(* IEC 61131-3 sources: daoli-st-library/DL_Process (part 30) *)

(* ---- FB_DL_DateCoderPosition.st ---- *)
(*==============================================================================
 * 组件名称 (Component)  : FB_DL_DateCoderPosition
 * 所属子库 (Sublibrary) : DL_Process
 * 当前版本 (Version)    : 1.0.0
 * 兼容性 (Platform)     : CODESYS 3.5+ / TwinCAT 3 / 汇川 InoProShop / 施耐德 Machine Expert
 *                         仅依赖 Standard.library（R_TRIG / ABS），零厂商私有库
 * 功能描述 (Function)   : 喷码日期位置偏移与缺失检测。检测触发沿按视觉检出
 *                         电平分派：未检出 → 缺失计数 + bMissing 锁存；检出
 *                         → 位置偏差 = 实测 - 期望，容差内 bPosOk，超差偏移
 *                         计数。判定结果锁存回放至下一触发沿（诊断资产）。
 *                         与 MarkPositionLatch（喷印位锁存）分工：本件是定
 *                         容差判偏移/缺失的诊断件。
 * 来源标签 (Origin)     : ROADMAP §21.4 R13 池（L907），自研 clean-room
 * 边界语义 (Boundary)   : ① 触发沿位置 NaN：按缺失域分派（视觉数据不可信 =
 *                         本拍无有效读码，归缺失语义安全侧）；
 *                         ② 容差/期望位置域闸 → 组态故障；
 *                         ③ 缺失/偏移计数 UDINT 独立成员（R190 归因唯一）；
 *                         ④ 状态锁存至下个触发沿（回放，不按当下输入重推断）。
 * 输出语义 (Fallback)   : 【R191】bEnable = FALSE → 判定出口冻结保持（诊断
 *                         资产）；eFault 相 → 冻结 + bError = TRUE。
 * 码位     (Codes)      : 按 R297 范式零 16# 码位硬编码；错误出口 BOOL+ENUM(eCause)。
 * 红线自检 (Redline)    : 7 项红线已自检：R1 零全局 ✓｜R2 零物理地址 ✓｜R3 纯 IEC ✓
 *                         R4 除零无涉/NaN 归缺失/组态闸 ✓｜R5 双语同行注释 ✓
 *                         R6 CASE 带 ELSE 兜底迁 eFault ✓｜R7 R_TRIG 段 0 无条件刷新 ✓
 * 验收向量 (Acceptance) : V1 期望 120.0、实测 121.4、容差 2.0 → 偏差 1.4，
 *                         bPosOk=TRUE；
 *                         V2 实测 124.0（偏差 4.0 超容差）→ nOffCnt+1，
 *                         bPosOk=FALSE；
 *                         V3 触发沿 bMarkPresent=FALSE → nMissCnt+1，
 *                         bMissing=TRUE。
 * 修订历史 (Revision)   : 2026-11-20  v1.0.0  R51 首版（批 3 · 序号 13）
 *==============================================================================*)
TYPE E_DL_DcpState :
(
    eIdle  := 0,                             (* 待使能 / Idle *)
    eInspect := 10,                          (* 检测运行 / Inspect run *)
    eFault := 90                             (* 故障锁存相 / Fault latched phase *)
);
END_TYPE

TYPE E_DL_DcpCause :
(
    eNone       := 0,                        (* 无故障成因 / No cause *)
    eCfgIllegal := 1,                        (* 组态非法：容差越域 / Illegal config *)
    ePhaseBad   := 2                         (* 非法相位兜底 / Illegal phase fallback *)
);
END_TYPE

FUNCTION_BLOCK FB_DL_DateCoderPosition
VAR_INPUT
    fMarkPos    : LREAL := 0.0;              (* 视觉测得喷码位置 [mm] / Measured mark position *)
    fMarkSp     : LREAL := 120.0;            (* 喷码期望位置，域 > 0 [mm] / Expected mark position *)
    fPosTol     : LREAL := 2.0;              (* 位置容差，域 > 0 [mm] / Position tolerance *)
    bMarkPresent: BOOL := FALSE;              (* 视觉检出电平 [-] / Vision present level *)
    bInspectTrig: BOOL := FALSE;             (* 检测触发电平（上升沿判定）[-] / Inspect trigger *)
    bEnable     : BOOL := TRUE;              (* 使能 [-] / Enable *)
    bReset      : BOOL := FALSE;             (* 复位命令，上升沿清全部 [-] / Reset command *)
END_VAR
VAR_OUTPUT
    fOffset     : LREAL;                     (* 位置偏差（实测 - 期望）[mm] / Position offset *)
    bPosOk      : BOOL;                      (* 位置合格判定（锁存回放）[-] / Position verdict *)
    bMissing    : BOOL;                      (* 喷码缺失锁存（下个触发沿或复位沿清）[-] / Missing latch *)
    nMissCnt    : UDINT;                     (* 缺失计数（独立成员，R190）[次] / Missing count *)
    nOffCnt     : UDINT;                     (* 偏移计数（独立成员，R190）[次] / Offset count *)
    nInspCnt    : UDINT;                     (* 累计检测次数 [次] / Inspect count *)
    eState      : E_DL_DcpState;             (* 状态出口 / State outlet *)
    eCause      : E_DL_DcpCause;             (* 故障成因出口 / Fault cause outlet *)
    bError      : BOOL;                      (* 故障锁存标志 [-] / Fault latch flag *)
END_VAR
VAR
    _eState   : E_DL_DcpState := E_DL_DcpState.eIdle;     (* 内部相位（CASE 唯一写入目标） / Internal phase *)
    _eCause   : E_DL_DcpCause := E_DL_DcpCause.eNone;     (* 故障成因锁存量 / Latched cause *)
    rtTrig    : R_TRIG;                      (* 触发沿实例，段 0 无条件调用 / Trigger edge instance *)
    rtReset   : R_TRIG;                      (* 复位沿实例，段 0 无条件调用 / Reset edge instance *)
    _fOff     : LREAL;                       (* 偏差派生量 [mm] / Offset derived *)
    _nMiss    : UDINT;                       (* 缺失计数锁存 [次] / Missing count latch *)
    _nOff     : UDINT;                       (* 偏移计数锁存 [次] / Offset count latch *)
    _nInsp    : UDINT;                       (* 检测计数锁存 [次] / Inspect count latch *)
    _bPosBad  : BOOL;                        (* 位置非有限当拍量 [-] / Non-finite position *)
    _bFault   : BOOL;                        (* 故障锁存位 / Latched fault bit *)
    _bCfgBad  : BOOL;                        (* 组态非法当拍量 / Illegal config this scan *)
END_VAR
VAR CONSTANT
    DL_DCP_EPS : LREAL := 1.0E-9;            (* 容差判零容差 [mm] / Tolerance epsilon *)
END_VAR

(* —— 段 0：当拍判据派生 + 沿实例无条件刷新（R228A） —— *)
_bCfgBad := (fPosTol <= DL_DCP_EPS) OR (fMarkSp <= 0.0);   (* 组态闸（R151 全引脚） / Config gate *)
rtTrig(CLK := bInspectTrig);                 (* 触发沿每拍必调 / Trigger edge every scan *)
rtReset(CLK := bReset);                      (* 复位沿每拍必调 / Reset edge every scan *)
_bPosBad := (fMarkPos <> fMarkPos) OR ((fMarkPos - fMarkPos) <> (fMarkPos - fMarkPos));   (* 位置 NaN 自反 + Inf 差判 / Non-finite position *)

(* —— 段 1：单拍量预清零（R107） —— *)
_fOff := 0.0;                                (* 偏差预清（判定拍内派生，R285） / Offset preset *)
bPosOk := FALSE;                             (* 判定预清（锁存拍内覆盖） / Verdict preset *)

(* —— 段 2：复位沿处理（作用域：清故障 + 清计数 + 清判定锁存 + 清出口 + 迁 eIdle，R283 逐项声明） —— *)
IF rtReset.Q THEN
    _bFault := FALSE;                        (* 清故障锁存 / Clear fault *)
    _eCause := E_DL_DcpCause.eNone;          (* 清成因 / Clear cause *)
    _nMiss := 0;                             (* 清缺失计数 / Clear miss count *)
    _nOff := 0;                              (* 清偏移计数 / Clear offset count *)
    _nInsp := 0;                             (* 清检测计数 / Clear inspect count *)
    bMissing := FALSE;                       (* 清缺失锁存（复位沿清除路径） / Clear missing latch *)
    bPosOk := FALSE;                         (* 清判定出口 / Clear verdict outlet *)
    fOffset := 0.0;                          (* 清偏差出口 / Clear offset outlet *)
    _eState := E_DL_DcpState.eIdle;          (* 迁待机相 / Back to idle *)
END_IF

(* —— 段 3：组态闸故障锁存（R45 配对；锁存至复位沿，R189） —— *)
IF _bCfgBad AND NOT _bFault THEN
    _bFault := TRUE;                         (* 锁存故障位 / Latch fault *)
    _eCause := E_DL_DcpCause.eCfgIllegal;    (* 成因：组态非法 / Cause: illegal config *)
    _eState := E_DL_DcpState.eFault;         (* 同步迁故障相 / Migrate to fault *)
END_IF

(* —— 段 4：CASE 主状态机（ELSE 兜底迁 eFault，红线 6） —— *)
CASE _eState OF
    E_DL_DcpState.eIdle:                     (* 待机相 / Idle *)
        IF bEnable AND NOT _bFault THEN
            _eState := E_DL_DcpState.eInspect;   (* 进入检测 / Enter inspect *)
        END_IF
    E_DL_DcpState.eInspect:                  (* 检测相：触发沿分派判定 / Inspect *)
        IF NOT bEnable THEN
            _eState := E_DL_DcpState.eIdle;  (* 失能回待机 / Back to idle *)
        ELSIF rtTrig.Q THEN                  (* 触发沿执行 / On trigger edge *)
            _nInsp := _nInsp + 1;            (* 检测计数（UDINT 回绕工程安全） / Count inspect *)
            IF (NOT bMarkPresent) OR _bPosBad THEN   (* 未检出或位置坏值：归缺失域（边界①安全侧） / Missing domain *)
                _nMiss := _nMiss + 1;        (* 缺失计数（独立成员） / Count missing *)
                bMissing := TRUE;            (* 缺失锁存（下个沿或复位清，边界④） / Latch missing *)
                bPosOk := FALSE;             (* 判定回放刷新 / Verdict replay *)
            ELSE
                _fOff := fMarkPos - fMarkSp; (* 偏差派生（减法无除零） / Offset derive *)
                fOffset := _fOff;            (* 偏差出口刷新 / Offset outlet *)
                IF ABS(_fOff) <= fPosTol THEN
                    bPosOk := TRUE;          (* 容差内合格 / In tolerance *)
                    bMissing := FALSE;       (* 检出合格拍清缺失锁存（触发沿清除路径，边界④） / Clear missing on pass *)
                ELSE
                    _nOff := _nOff + 1;      (* 偏移计数（独立成员） / Count offset *)
                    bPosOk := FALSE;         (* 超差不合格 / Out of tolerance *)
                END_IF
            END_IF
        END_IF                               (* 非触发拍：状态锁存回放（边界④） / Replay between edges *)
    E_DL_DcpState.eFault:                    (* 故障相：冻结保持，仅复位沿出 / Fault *)
        ;                                    (* 锁存回放（R28） / Replay from latch *)
    ELSE                                     (* 非法相位兜底迁安全态 / Illegal phase fallback *)
        _eState := E_DL_DcpState.eFault;     (* 迁故障相 / To fault *)
        _bFault := TRUE;                     (* 同步锁存 / Latch *)
        _eCause := E_DL_DcpCause.ePhaseBad;  (* 成因：非法相位 / Cause: illegal phase *)
END_CASE

(* —— 段 5：出口映射（bError/eState 同源，R191） —— *)
nMissCnt := _nMiss;                          (* 缺失计数出口 / Miss outlet *)
nOffCnt := _nOff;                            (* 偏移计数出口 / Offset outlet *)
nInspCnt := _nInsp;                          (* 检测计数出口 / Inspect outlet *)
bError := _bFault;                           (* 故障标志镜像 / Fault flag mirror *)
eState := _eState;                           (* 状态出口 / State outlet *)
eCause := _eCause;                           (* 成因出口 / Cause outlet *)
END_FUNCTION_BLOCK

(* ---- FB_DL_DesiccantRegenSeq.st ---- *)
(*
  组件名 Component   : FB_DL_DesiccantRegenSeq
  子库 Sublibrary    : DL_Process
  版本 Version       : 1.0.0
  兼容性 Platform    : CODESYS 3.5 / TwinCAT 3 / 汇川 InoProShop / Machine Expert（仅 Standard.library）
  功能 Function      : 干燥剂吸附塔再生顺控（ISA-88 相语义最小子集）：
                       1) 四相顺控：吸附（eAdsorb）→ 再生（eRegen）→ 吹冷（eCool）→
                       切换驻留（eSwitchDwell）→ 回吸附，吸附时长由 tAdsorbDur 承载；
                       2) 塔间轮换：A/B 双塔，eSwitchDwell 相完成阀组切换并翻转
                       bTowerAActive/bTowerBActive（切换指令单点出口）；
                       3) 再生温度曲线监视：再生相内再生温度须在
                       [fRegenTempLoC, fRegenTempHiC] 曲线带内，越带持续 tTempDevTo
                       → 故障锁存；
                       4) 各相计时独立 TON 实例（禁跨相复用，R228A）。
  边界 Boundary      : ① 本件只出阀组/加热指令与塔选通，不写物理 IO；
                       ② 吹冷相退出双条件：吹冷计时到 或 出口温度低于 fCoolEndC
                       （事件达成 + 前置消失双路径）；再生许可不满足时吸附相驻留等待；
                       ③ 故障锁存解除唯一路径 = bReset 上升沿（输入引脚，恒可达）；
                       ④ 无全局变量引用、无外部变量声明、无物理地址寻址。
  依赖 Depends       : Standard.library（R_TRIG / TON）
  溯源 Origin        : 道莅自研 clean-room（参考 t2-8-isa88 相语义分类与参数域，
                       零代码行复制）
  码位 Code          : 16#06_0_BE（Process 段 0006，B 子带 BE 格）
  码表 Error codes（本件格 06_0_BE，单轨子道：故障 0x02BE / 信息 0x01BE）:
    16#0006_02BE 故障级：再生顺控故障总码（再生温度越带 / 切换超时 / 组态非法 /
                 输入非有限），锁存至复位
    16#0006_01BE 信息级：塔切换完成沿（eSwitchDwell → eAdsorb 迁移拍）
  修订历史 Revision  :
    2026-11-19  v1.0.0  R44 首版（批次 3 · 序号 15）
*)

TYPE E_DL_DrsPhase :
(
    eIdle        := 0,   // 空闲：未使能 / Idle, not enabled
    eAdsorb      := 10,  // 吸附：当前塔吸附运行 / Adsorbing on active tower
    eRegen       := 20,  // 再生：离线塔再生加热 / Regenerating offline tower
    eCool        := 30,  // 吹冷：再生塔吹冷 / Cooling regenerated tower
    eSwitchDwell := 40,  // 切换：塔间阀组切换驻留 / Switching towers dwell
    eFault       := 90   // 故障：总码锁存 / Fault, latched
);
END_TYPE

FUNCTION_BLOCK FB_DL_DesiccantRegenSeq
VAR_INPUT
    bEnable      : BOOL;                   // 使能（电平）[-] / Enable
    bReset       : BOOL;                   // 上升沿清故障锁存 [-] / Reset edge
    bRegenPermissive: BOOL;                // 再生许可（电平）[-] / Regen permissive
    fRegenTempC  : REAL;                   // 再生温度 [摄氏度] / Regen temperature
    fCoolOutTempC: REAL;                   // 吹冷出口温度 [摄氏度] / Cooling outlet temperature
    tAdsorbDur   : TIME := T#8H;           // 吸附时长 [毫秒] / Adsorption duration
    tRegenDur    : TIME := T#4H;           // 再生时长 [毫秒] / Regen duration
    tCoolMaxDur  : TIME := T#2H;           // 吹冷最大时长 [毫秒] / Cooling max duration
    tSwitchDur   : TIME := T#60S;          // 切换驻留 [毫秒] / Switch dwell
    fRegenTempLoC: REAL := 120.0;          // 再生温度带下限 [摄氏度] / Regen band floor
    fRegenTempHiC: REAL := 200.0;          // 再生温度带上限 [摄氏度] / Regen band ceiling
    fCoolEndC    : REAL := 45.0;           // 吹冷结束温度 [摄氏度] / Cooling end temperature
    tTempDevTo   : TIME := T#30S;          // 温度越带确认窗 [毫秒] / Temperature deviation timeout
END_VAR
VAR_OUTPUT
    bTowerAActive: BOOL;                   // A 塔吸附选通 [-] / Tower A active
    bTowerBActive: BOOL;                   // B 塔吸附选通 [-] / Tower B active
    bRegenHeatCmd: BOOL;                   // 再生加热指令 [-] / Regen heat command
    bRegenCoolCmd: BOOL;                   // 吹冷指令 [-] / Regen cool command
    bSwitchCmd   : BOOL;                   // 塔切换指令（驻留相电平）[-] / Tower switch command
    ePhase       : E_DL_DrsPhase;          // 相位出口，段尾单点映射 / Phase outlet
    bError       : BOOL;                   // 故障锁存标志 [-] / Fault latch flag
    uErrId       : UDINT;                  // 事件码，0 = 无事件 / Event code
END_VAR
VAR
    rtReset   : R_TRIG;                    // 复位沿实例，段 0 无条件刷新 / Reset edge
    tonAdsorb : TON;                       // 吸附计时（独立实例） / Adsorption timer
    tonRegen  : TON;                       // 再生计时（独立实例） / Regen timer
    tonCoolMax: TON;                       // 吹冷最大计时（独立实例） / Cooling max timer
    tonSwitch : TON;                       // 切换驻留计时（独立实例） / Switch dwell timer
    tonTempDevTo: TON;                     // 温度越带确认（专用超时件命名） / Temp deviation timeout
    _ePhase   : E_DL_DrsPhase := E_DL_DrsPhase.eIdle;  // 内部相位（CASE 唯一写入目标）/ Internal phase
    _bTowerA  : BOOL := TRUE;              // 内部塔选（TRUE = A 塔吸附）/ Internal tower select
    _bFault   : BOOL;                      // 故障锁存位（锁存量） / Latched fault bit
    _uFault   : UDINT;                     // 故障码锁存（锁存量） / Latched fault code
    _bCfgBad  : BOOL;                      // 组态非法当拍量 [-] / Config illegal flag
    _bNonFin  : BOOL;                      // 输入非有限当拍量 [-] / Non-finite input flag
    _bTempDev : BOOL;                      // 温度越带当拍量 [-] / Temperature deviation flag
END_VAR
VAR CONSTANT
    DL_ABS_MAX : REAL := 1.0E30;           // 有限值判定上界 [摄氏度] / Finite bound
    DL_ZERO    : REAL := 0.0;              // 零常量 [摄氏度] / Zero constant
END_VAR

(* —— 段 0｜沿与定时器每拍无条件刷新（禁置于 IF/CASE 内；各相独立实例禁复用） —— *)
rtReset(CLK := bReset);
tonAdsorb (IN := (_ePhase = E_DL_DrsPhase.eAdsorb) AND (NOT _bFault), PT := tAdsorbDur);
tonRegen  (IN := (_ePhase = E_DL_DrsPhase.eRegen) AND (NOT _bFault), PT := tRegenDur);
tonCoolMax(IN := (_ePhase = E_DL_DrsPhase.eCool) AND (NOT _bFault), PT := tCoolMaxDur);
tonSwitch (IN := (_ePhase = E_DL_DrsPhase.eSwitchDwell) AND (NOT _bFault), PT := tSwitchDur);
_bTempDev := (_ePhase = E_DL_DrsPhase.eRegen)
             AND ((fRegenTempC < fRegenTempLoC) OR (fRegenTempC > fRegenTempHiC));
tonTempDevTo(IN := _bTempDev AND (NOT _bFault), PT := tTempDevTo);

(* —— 段 1｜瞬时量预清零（锁存量 _bFault/_uFault/_bTowerA 不入清单） —— *)
uErrId   := 16#0000_0000;
_bCfgBad := FALSE;
_bNonFin := FALSE;

(* —— 段 2｜复位沿：故障一次性清干净，相位回空闲 —— *)
IF rtReset.Q THEN
    _bFault := FALSE;
    _uFault := 16#0000_0000;
    _ePhase := E_DL_DrsPhase.eIdle;
END_IF

(* —— 段 3｜组态闸与非有限判据（覆盖全部参与判据换算引脚） —— *)
IF (fRegenTempLoC >= fRegenTempHiC) OR (tAdsorbDur = T#0S) OR (tRegenDur = T#0S)
   OR (tCoolMaxDur = T#0S) OR (tSwitchDur = T#0S) OR (tTempDevTo = T#0S) THEN
    _bCfgBad := TRUE;
END_IF
IF (fRegenTempC <> fRegenTempC) OR ((fRegenTempC - fRegenTempC) <> DL_ZERO)
   OR (fCoolOutTempC <> fCoolOutTempC) OR ((fCoolOutTempC - fCoolOutTempC) <> DL_ZERO) THEN
    _bNonFin := TRUE;
END_IF

(* —— 段 4｜主状态机：六态全覆盖 + ELSE 兜底 —— *)
CASE _ePhase OF

E_DL_DrsPhase.eIdle:
    bTowerAActive := FALSE;
    bTowerBActive := FALSE;
    bRegenHeatCmd := FALSE;
    bRegenCoolCmd := FALSE;
    bSwitchCmd    := FALSE;
    IF bEnable AND (NOT _bCfgBad) THEN
        _bTowerA := TRUE;                // 入运行相：A 塔先吸附（固定初序）
        _ePhase  := E_DL_DrsPhase.eAdsorb;
    ELSIF bEnable AND _bCfgBad THEN
        _bFault := TRUE;
        _uFault := 16#0006_02BE;
        bError  := TRUE;
        _ePhase := E_DL_DrsPhase.eFault;
    END_IF

E_DL_DrsPhase.eAdsorb:
    bTowerAActive := _bTowerA;
    bTowerBActive := NOT _bTowerA;
    bRegenHeatCmd := FALSE;
    bRegenCoolCmd := FALSE;
    bSwitchCmd    := FALSE;
    IF _bNonFin THEN
        _bFault := TRUE;
        _uFault := 16#0006_02BE;
        bError  := TRUE;
        _ePhase := E_DL_DrsPhase.eFault;
    ELSIF NOT bEnable THEN
        _ePhase := E_DL_DrsPhase.eIdle;  // 使能撤销回空闲
    ELSIF tonAdsorb.Q AND bRegenPermissive THEN
        _ePhase := E_DL_DrsPhase.eRegen; // 吸附时长到且再生许可满足：进再生
    ELSIF tonAdsorb.Q THEN
        ;                                // 吸附时长到但许可未满足：吸附相驻留等待（退出前置消失路径）
    END_IF

E_DL_DrsPhase.eRegen:
    bTowerAActive := _bTowerA;
    bTowerBActive := NOT _bTowerA;
    bRegenHeatCmd := TRUE;
    bRegenCoolCmd := FALSE;
    bSwitchCmd    := FALSE;
    IF _bNonFin OR tonTempDevTo.Q THEN
        _bFault := TRUE;                 // 温度越带或输入非法：锁存
        _uFault := 16#0006_02BE;
        bError  := TRUE;
        _ePhase := E_DL_DrsPhase.eFault;
    ELSIF NOT bEnable THEN
        _ePhase := E_DL_DrsPhase.eIdle;  // 使能撤销回空闲
    ELSIF tonRegen.Q THEN
        _ePhase := E_DL_DrsPhase.eCool;  // 迁出条件 1：再生时长到
    END_IF

E_DL_DrsPhase.eCool:
    bTowerAActive := _bTowerA;
    bTowerBActive := NOT _bTowerA;
    bRegenHeatCmd := FALSE;
    bRegenCoolCmd := TRUE;
    bSwitchCmd    := FALSE;
    IF _bNonFin THEN
        _bFault := TRUE;
        _uFault := 16#0006_02BE;
        bError  := TRUE;
        _ePhase := E_DL_DrsPhase.eFault;
    ELSIF NOT bEnable THEN
        _ePhase := E_DL_DrsPhase.eIdle;  // 使能撤销回空闲
    ELSIF (fCoolOutTempC <= fCoolEndC) OR tonCoolMax.Q THEN
        _ePhase := E_DL_DrsPhase.eSwitchDwell;   // 迁出双条件：温度达成 或 吹冷计时到
    END_IF

E_DL_DrsPhase.eSwitchDwell:
    bTowerAActive := FALSE;
    bTowerBActive := FALSE;
    bRegenHeatCmd := FALSE;
    bRegenCoolCmd := FALSE;
    bSwitchCmd    := TRUE;               // 切换指令（驻留相电平）
    IF _bNonFin THEN
        _bFault := TRUE;
        _uFault := 16#0006_02BE;
        bError  := TRUE;
        _ePhase := E_DL_DrsPhase.eFault;
    ELSIF NOT bEnable THEN
        _ePhase := E_DL_DrsPhase.eIdle;  // 使能撤销回空闲
    ELSIF tonSwitch.Q THEN
        _bTowerA := NOT _bTowerA;        // 塔间轮换翻转
        uErrId := 16#0006_01BE;          // 信息级：塔切换完成沿
        _ePhase := E_DL_DrsPhase.eAdsorb;    // 回吸附相（待机可返回路径）
    END_IF

E_DL_DrsPhase.eFault:
    bTowerAActive := FALSE;
    bTowerBActive := FALSE;
    bRegenHeatCmd := FALSE;              // 故障相：加热指令安全侧撤销
    bRegenCoolCmd := FALSE;
    bSwitchCmd    := FALSE;
    bError := TRUE;
    ;                                    // 故障相驻留：只认复位沿（段 2 迁出）

ELSE
    _bFault := TRUE;                     // 兜底：非法相位锁存
    _uFault := 16#0006_02BE;
    bError  := TRUE;
    _ePhase := E_DL_DrsPhase.eFault;
END_CASE

(* —— 段 5｜相位出口单点映射 —— *)
ePhase := _ePhase;
END_FUNCTION_BLOCK

(* ---- FB_DL_DieBinCounter.st ---- *)
(*
  Name        : FB_DL_DieBinCounter
  Category    : DL_Process
  Version     : 1.0.0
  Purpose     : 晶粒分箱计数与满箱切换：按来料脉冲累加晶粒数，接近容量即预警，满箱置切换请求，收到换箱确认后清零并箱号递增；/ Count dies per bin with near-full warning, full-bin switch request and post-acknowledge bin index advance
  溯源        : ROADMAP L647（未勾真缺口），IEC 61131-3 标准语义的道莅防御性实现
  Boundary    : ① 组态闸：箱容量 < 2 / 预警余量 < 0 或 >= 容量 → 锁存故障（余量需严格小于容量，否则预警永不触发）；
                ② 计数只认单拍脉冲上升沿（防电平长时间为真时多计）；
                ③ 满箱锁存后不再接收计数脉冲（拒收计 nReject），避免溢出把计数推过容量；
                ④ 切换请求为状态量（eFull 相保持），换箱确认为上升沿（跨周期动作不用单拍标志门控）；
                ⑤ 箱号 UDINT 饱和累加，满容量计数上限钳到箱容量（防越界显示）。
*)
TYPE E_DL_DbcState :
(
    eIdle   := 0,                            (* 未使能 / Disabled *)
    eCount  := 10,                           (* 计数中 / Counting *)
    eFull   := 20,                           (* 满箱待换箱 / Full, awaiting switch *)
    eFault  := 90                            (* 故障锁存相 / Fault latched *)
);
END_TYPE

TYPE E_DL_DbcCause :
(
    eNone       := 0,                        (* 无故障成因 / No cause *)
    eCfgIllegal := 1,                        (* 组态非法：容量/余量越域 / Illegal config *)
    ePhaseBad   := 2                         (* 非法相位兜底 / Illegal phase fallback *)
);
END_TYPE

FUNCTION_BLOCK FB_DL_DieBinCounter
VAR_INPUT
    bDiePulse   : BOOL := FALSE;             (* 晶粒来料脉冲（上升沿计 1 颗）[-] / Die arrival pulse, rising edge counts one *)
    nBinCap     : INT := 5000;               (* 箱容量，域 >= 2 [颗] / Bin capacity, >= 2 *)
    nWarnMargin : INT := 200;                (* 满箱预警余量，域 0 <= x < nBinCap [颗] / Near-full margin *)
    bSwitchAck  : BOOL := FALSE;             (* 换箱完成确认（上升沿）[-] / Bin switch acknowledge edge *)
    bEnable     : BOOL := TRUE;              (* 使能 [-] / Enable *)
    bReset      : BOOL := FALSE;             (* 复位命令，上升沿清计数/箱号/故障 [-] / Reset command *)
END_VAR
VAR_OUTPUT
    nCount      : INT;                       (* 当前箱已装颗数（钳到容量）[颗] / Current bin count, clamped to capacity *)
    nBinIdx     : UDINT;                     (* 当前箱号（从 1 起，饱和）[-] / Current bin index, from 1, saturated *)
    bNearFull   : BOOL;                      (* 接近满箱预警 [-] / Near-full warning *)
    bBinFull    : BOOL;                      (* 满箱锁存 [-] / Bin full latch *)
    bSwitchReq  : BOOL;                      (* 换箱请求（满箱相保持）[-] / Switch request while full *)
    nReject     : INT;                       (* 满箱期拒收脉冲数（诊断，饱和）[颗] / Rejected pulses while full *)
    eState      : E_DL_DbcState;             (* 状态出口 / State outlet *)
    eCause      : E_DL_DbcCause;             (* 故障成因出口（R190 归因唯一） / Fault cause outlet *)
    bError      : BOOL;                      (* 故障锁存标志 [-] / Fault latch flag *)
END_VAR
VAR
    _eState  : E_DL_DbcState := E_DL_DbcState.eIdle;     (* 内部相位（CASE 唯一写入目标） / Internal phase *)
    _eCause  : E_DL_DbcCause := E_DL_DbcCause.eNone;     (* 故障成因锁存量 / Latched cause *)
    rtPulse  : R_TRIG;                       (* 来料脉冲上升沿，段 0 无条件调用 / Die pulse edge *)
    rtAck    : R_TRIG;                       (* 换箱确认上升沿，段 0 无条件调用 / Ack edge *)
    rtReset  : R_TRIG;                       (* 复位沿实例，段 0 无条件调用 / Reset edge *)
    _bFault  : BOOL;                         (* 故障锁存位 / Latched fault bit *)
    _bCfgBad : BOOL;                         (* 组态非法当拍量 / Illegal config this scan *)
    _bFull   : BOOL;                         (* 满箱锁存位 / Full latch *)
    _nCount  : INT;                          (* 计数内部量 [颗] / Count internal *)
    _nRej    : INT;                          (* 拒收计数内部量 [颗] / Reject internal *)
    _nWarnTh : INT;                          (* 预警门槛 = 容量 - 余量 [颗] / Warning threshold *)
END_VAR
VAR CONSTANT
    DL_DBC_CNTMAX : UDINT := 4294967295;     (* 箱号饱和上限（R28）[-] / Bin index cap *)
    DL_DBC_REJMAX : INT   := 32767;          (* 拒收计数饱和上限（INT 可表上限）[颗] / Reject count cap *)
    DL_DBC_NMIN   : INT   := 2;              (* 容量下限（需能容纳预警余量逻辑）[颗] / Capacity lower bound *)
END_VAR

(* —— 段 0：当拍判据派生 + 实例无条件刷新（R228A） —— *)
_bCfgBad := (nBinCap < DL_DBC_NMIN)                                            (* 容量域闸 / Capacity gate *)
            OR (nWarnMargin < 0) OR (nWarnMargin >= nBinCap);                  (* 余量域闸（须严格小于容量） / Margin gate *)
rtPulse(CLK := bDiePulse);                                                     (* 来料沿每拍必调 / Pulse edge every scan *)
rtAck(CLK := bSwitchAck);                                                      (* 确认沿每拍必调 / Ack edge every scan *)
rtReset(CLK := bReset);                                                        (* 复位沿每拍必调 / Reset edge every scan *)
_nWarnTh := nBinCap - nWarnMargin;                                             (* 预警门槛反算（容量 > 余量，差恒正）[颗] / Warning threshold *)

(* —— 段 1：单拍量预清零（R107） —— *)
bNearFull := FALSE;                                                            (* 预警位预清 / Near-full preset *)
bSwitchReq := FALSE;                                                           (* 换箱请求预清（仅满箱相置位） / Request preset *)

(* —— 段 2：复位沿处理（作用域：清故障 + 清计数 + 清箱号 + 清满箱锁存 + 迁 eIdle，R283 逐项声明） —— *)
IF rtReset.Q THEN
    _bFault := FALSE;                                                          (* 清故障锁存 / Clear fault *)
    _eCause := E_DL_DbcCause.eNone;                                            (* 清成因 / Clear cause *)
    _bFull := FALSE;                                                           (* 清满箱锁存（隐性回夹防护） / Clear full latch *)
    _nCount := 0;                                                              (* 清计数 / Clear count *)
    _nRej := 0;                                                                (* 清拒收计数 / Clear reject count *)
    nCount := 0;                                                               (* 清计数出口 / Clear count outlet *)
    nBinIdx := 1;                                                              (* 箱号回 1（从 1 起） / Bin index back to 1 *)
    bBinFull := FALSE;                                                         (* 清满箱出口 / Clear full outlet *)
    nReject := 0;                                                              (* 清拒收出口 / Clear reject outlet *)
    _eState := E_DL_DbcState.eIdle;                                            (* 迁未使能相 / Back to idle *)
END_IF

(* —— 段 3：组态故障锁存（锁存至复位沿，R189） —— *)
IF _bCfgBad AND NOT _bFault THEN
    _bFault := TRUE;                                                           (* 锁存故障位 / Latch fault *)
    _eCause := E_DL_DbcCause.eCfgIllegal;                                      (* 成因：组态非法 / Cause: illegal config *)
    _eState := E_DL_DbcState.eFault;                                           (* 同步迁故障相 / Migrate to fault *)
END_IF

(* —— 段 4：CASE 主状态机（ELSE 兜底迁 eFault，红线 6） —— *)
CASE _eState OF
    E_DL_DbcState.eIdle:                                                       (* 未使能：不计数 / Disabled *)
        nCount := _nCount;                                                     (* 出口镜像（保留进度） / Outlet mirror *)
        IF bEnable AND NOT _bFault THEN
            IF nBinIdx = 0 THEN
                nBinIdx := 1;                                                  (* 未初始化箱号兜底为 1（首次使能） / Init bin index *)
            END_IF
            _eState := E_DL_DbcState.eCount;                                   (* 使能进入计数 / Enter counting *)
        END_IF
    E_DL_DbcState.eCount:                                                      (* 计数相：脉冲累加 + 满箱推进 / Counting *)
        IF NOT bEnable THEN
            _eState := E_DL_DbcState.eIdle;                                    (* 失能回未使能 / Back to idle *)
        ELSE
            IF rtPulse.Q THEN                                                  (* 单拍脉冲上升沿计 1 颗 / One die per rising edge *)
                IF _nCount < nBinCap THEN
                    _nCount := _nCount + 1;                                    (* 容量内递增（满后拒收） / Increment within capacity *)
                END_IF
            END_IF
            IF _nCount >= nBinCap THEN
                _nCount := nBinCap;                                            (* 计数钳到容量（防越界显示） / Clamp to capacity *)
                _bFull := TRUE;                                                (* 满箱锁存 / Latch full *)
            END_IF
            nCount := _nCount;                                                 (* 计数出口 / Count outlet *)
            IF NOT _bFull THEN
                IF _nCount >= _nWarnTh THEN
                    bNearFull := TRUE;                                         (* 接近满箱预警 / Near-full warning *)
                END_IF
            END_IF
            bBinFull := _bFull;                                                (* 满箱出口镜像（名实同源，R191） / Full outlet mirror *)
            IF _bFull THEN
                _eState := E_DL_DbcState.eFull;                                (* 迁满箱相（请求换箱） / To full *)
            END_IF
        END_IF
    E_DL_DbcState.eFull:                                                       (* 满箱相：保持请求，拒收脉冲，等确认 / Full *)
        bBinFull := TRUE;                                                      (* 满箱出口保持 / Full outlet held *)
        bSwitchReq := TRUE;                                                    (* 换箱请求状态量保持（非单拍标志） / Request held as state *)
        nCount := _nCount;                                                     (* 计数出口保持 / Count outlet held *)
        IF rtPulse.Q THEN
            IF _nRej < DL_DBC_REJMAX THEN
                _nRej := _nRej + 1;                                            (* 满箱期拒收脉冲计数（诊断） / Count rejects *)
            END_IF
        END_IF
        nReject := _nRej;                                                      (* 拒收出口 / Reject outlet *)
        IF rtAck.Q THEN                                                        (* 换箱确认上升沿：清零换箱 / Ack: reset bin *)
            _nCount := 0;                                                      (* 清计数 / Clear count *)
            _bFull := FALSE;                                                   (* 清满箱锁存 / Clear full *)
            bBinFull := FALSE;                                                 (* 清满箱出口 / Clear full outlet *)
            nCount := 0;                                                       (* 清计数出口 / Clear count outlet *)
            IF nBinIdx < DL_DBC_CNTMAX THEN
                nBinIdx := nBinIdx + 1;                                        (* 箱号饱和递增 / Saturating bin index *)
            END_IF
            _eState := E_DL_DbcState.eCount;                                   (* 回计数相 / Back to counting *)
        END_IF
    E_DL_DbcState.eFault:                                                      (* 故障相：冻结保持末值，仅复位沿出 / Fault *)
        ;                                                                      (* 锁存回放（R28） / Replay from latch *)
    ELSE                                                                       (* 非法相位兜底迁安全态 / Illegal phase fallback *)
        _eState := E_DL_DbcState.eFault;                                       (* 迁故障相 / To fault *)
        _bFault := TRUE;                                                       (* 同步锁存 / Latch *)
        _eCause := E_DL_DbcCause.ePhaseBad;                                    (* 成因：非法相位 / Cause: illegal phase *)
END_CASE

(* —— 段 5：出口映射（bError/eState 同源，R191） —— *)
bError := _bFault;                                                             (* 故障标志镜像 / Fault flag mirror *)
eState := _eState;                                                             (* 状态出口 / State outlet *)
eCause := _eCause;                                                             (* 成因出口 / Cause outlet *)
END_FUNCTION_BLOCK

(* ---- FB_DL_DowntimeClassifier.st ---- *)
(*
    FB_DL_DowntimeClassifier —— 停机原因自动分类
    ------------------------------------------------------------------
    分类      : DL_Process / Oee
    前缀      : FB_DL_
    版本      : 1.0.0
    溯源      : T2-7 PackML / OMAC（只借「停机原因 / 未计划停机归因」的公开语义分类，
                不做 17 态全集——全集唯一属主是 FB_DL_PackMlStateMachine）；
                时长口径、计数口径、仲裁与码位 100% 自有；clean-room 重写，
                未复制任何闭源厂商源码，参考实现仅限 MIT/Apache 许可
    平台      : 纯 IEC 61131-3，CODESYS V3.5+ / TwinCAT 3 / InoProShop 通用
    作者      : 道莅代码库 · PLC编程专家（R18）
    ------------------------------------------------------------------
    功能说明  : 设备停转时自动抓取「哪个原因源先动」，给出停机原因序号与停机时长；
                同拍多源按序号最小仲裁（索引最小即优先级最高），超时未归类标未分类；
                三道防御：时间参数自相矛盾闸（最短时长大于归类等待上限即统计不可信）
                → 时长累加前先钳位（TIME 加法溢出在三平台行为不同，必须先比后加）
                → 计数饱和闸（UDINT 回绕会让台账出现天文数字）；
                结算纪律：只在停机结束那一拍累加时长与次数，停机中累加会重复计数；
                职责边界：刻意不做 OEE 三因子，该职责唯一属主是 FB_DL_OeeCalculator，
                避免两套统计口径打架。
    错误码    : 16#0005_01D2 同拍多源停机，已按源序号最小仲裁——信息级，不置故障
                16#0005_01D3 预留禁用（信息级，不得挪用）
                16#0005_02FF 停机超归类等待上限仍无原因源，判未分类（需人工补录）——故障级，需人工介入
                16#0005_0300 时间参数自相矛盾（归类上限小于最短时长或不为正）——故障级，统计冻结
                16#0005_0301 状态机落 ELSE 兜底（非法状态，回空闲）——故障级，回安全态
    码位总账  : 16#0005_01D2 用 / 16#0005_01D3 预留 ｜ 16#0005_02FF 用 / 16#0005_0300 用 / 16#0005_0301 用
    状态机    : E_DL_DowntimeState（eIdle / eStopped / eClassifying / eFault），
                CASE 含 ELSE 兜底，兜底固定置 eFault 与 0301
    采样约定  : 两个 TON 与三个 R_TRIG 在本体首部无条件调用；tMinDuration 与
                tMaxClassify 由工艺给定，改动后需一次复位使统计口径重新起算。
    修订记录  : 2026-11-16 v1.0.0 首次入库（R18）
*)

(*-----------------------------------------------------------------------------
 * 枚举: E_DL_DowntimeState（归属本功能块，与其同文件发布）
 * 含义: 停机归因状态机离散态，步长 10 留空位，故障态取 99 排末位
 *----------------------------------------------------------------------------*)
TYPE E_DL_DowntimeState :
(
    eIdle        := 0,   // 空闲：设备运行中，无停机在统计 / Idle, the machine runs and no downtime is being tracked
    eStopped     := 10,  // 停机中：尚未达到最短停机时长，随时可能被过滤 / Stopped, the minimum duration is not reached yet and may still be filtered out
    eClassifying := 20,  // 归类中：已超最短时长，等待原因源或归类上限 / Classifying, past the minimum duration, waiting for a cause or the classify limit
    eFault       := 99   // 故障：参数矛盾或非法状态，统计冻结 / Fault, contradictory parameters or an illegal state, statistics frozen
) UINT;
END_TYPE

FUNCTION_BLOCK FB_DL_DowntimeClassifier
VAR_INPUT
    bEnable          : BOOL;                   // 使能，FALSE 冻结统计（不清已累计值）/ enable, FALSE freezes the statistics without clearing them
    bReset           : BOOL;                   // 上升沿清累计与当前停机 / rising edge clears the totals and the current downtime
    bMachineRunning  : BOOL := FALSE;          // 设备运行信号，FALSE 且持续超最短时长即判停机 / machine running signal, FALSE beyond the minimum duration counts as downtime
    aStopCause       : ARRAY[0..7] OF BOOL;    // 8 路停机原因源，索引即优先级 0 最高 / 8 stop cause sources, the index is the priority, 0 highest
    tMinDuration     : TIME := T#5S;           // 最短停机时长，短于此不计入 [ms]，范围 100~600000 / minimum downtime filtered out below it [ms], range 100~600000
    tMaxClassify     : TIME := T#120S;         // 归类等待上限，超过仍无源即未分类 [ms] / classify wait limit, no source beyond it means unclassified [ms]
END_VAR
VAR_OUTPUT
    bDowntime     : BOOL;                      // 当前处于停机且已计时 / currently stopped and being timed
    tDownElapsed  : TIME;                      // 本次停机已持续时长 [ms] / elapsed time of the current downtime [ms]
    uActiveCause  : UINT;                      // 当前原因序号 0~7，16#FFFF = 未知 / current cause index 0~7, 16#FFFF = unknown
    uLastCause    : UINT;                      // 上次停机最终归因 / final cause of the previous downtime
    bUnclassified : BOOL;                      // 本次停机未归类（超上限或无源）/ the current downtime is unclassified
    auCauseCount  : ARRAY[0..7] OF UDINT;      // 各原因累计次数，饱和计数 [次] / accumulated count per cause, saturating [times]
    auCauseTime   : ARRAY[0..7] OF TIME;       // 各原因累计停机时长，饱和累加 [ms] / accumulated downtime per cause, saturating [ms]
    eErr          : UDINT;                     // 错误码，0=正常 / error id, 0=ok
    bError        : BOOL;                      // 故障标志，eErr 为故障级时 TRUE / error flag, TRUE on fault-level eErr
END_VAR
VAR
    fbTrigReset  : R_TRIG;                     // 复位沿检测实例，本体首部无条件刷新 / reset edge instance, refreshed unconditionally
    fbTrigRunOff : R_TRIG;                     // 运行信号下降沿实例 / running signal falling edge instance
    fbTrigRunOn  : R_TRIG;                     // 运行信号上升沿实例 / running signal rising edge instance
    fbMinDown    : TON;                        // 停机时长定时器，本体首部无条件刷新 / downtime duration timer, refreshed unconditionally
    fbClassify   : TON;                        // 归类等待定时器，本体首部无条件刷新 / classify wait timer, refreshed unconditionally
    eState       : E_DL_DowntimeState := E_DL_DowntimeState.eIdle; // 内部状态机步序 / internal state machine step
    uIdx         : UINT;                       // 原因源扫描游标 [路] / cause scan cursor [ch]
    uActCnt      : UINT;                       // 本拍有效原因源计数 [路] / active cause count this cycle [ch]
    bAnyCause    : BOOL;                       // 本拍存在原因源标志 / any cause active this cycle
    uFirstFound  : UINT;                       // 本拍首个为真的原因序号 / first active cause index this cycle
    uCauseCur    : UINT;                       // 本次停机已锁定的原因序号 / cause index locked for the current downtime
    tAccum       : TIME;                       // 单次停机时长累加中间量 [ms] / single downtime accumulation intermediate [ms]
    tClamped     : TIME;                       // 钳位中间量 [ms] / clamping intermediate [ms]
    bInit        : BOOL := FALSE;              // 首扫标志，初值 FALSE，判据 NOT bInit / first-scan flag, initial FALSE, tested with NOT
    bParamBad    : BOOL;                       // 时间参数矛盾标志 / contradictory time parameter flag
END_VAR
VAR CONSTANT
    DL_DTC_SRC_MAX  : UINT := 8;               // 原因源上限 [路] / cause source upper bound [ch]
    DL_DTC_NONE     : UINT := 16#FFFF;         // 未知原因哨兵 [无量纲] / unknown cause sentinel [dimensionless]
    DL_DTC_TIME_MAX : TIME := T#24H;           // 单次停机时长饱和值，防累加溢出 [ms] / single downtime saturation value against accumulation overflow [ms]
    DL_DTC_MAX_LOOP : UINT := 8;               // 循环守卫上限 [次] / loop guard upper limit [times]
    DL_DTC_MIN_DUR  : TIME := T#100MS;         // 最短停机时长下限 [ms] / minimum downtime lower bound [ms]
    DL_DTC_CNT_MAX  : UDINT := 16#FFFF_FFFE;   // 计数饱和值 [次] / count saturation value [times]
END_VAR

// 段 0｜输出与错误状态预置 / segment 0, preset outputs and error status
eErr := 0;                                     // 预置无错误 / preset no error
bError := FALSE;                               // 预置无故障 / preset no fault
bDowntime := FALSE;                            // 预置非停机 / preset not stopped
bUnclassified := FALSE;                        // 预置未判未分类 / preset not unclassified
bParamBad := FALSE;                            // 预置参数合法 / preset parameters valid
uActCnt := 0;                                  // 原因计数清零 / clear the cause count
bAnyCause := FALSE;                            // 原因标志清零 / clear the cause flag
uFirstFound := DL_DTC_NONE;                    // 首个原因先置哨兵 / the first cause starts at the sentinel

// 段 1｜时间参数闸：自相矛盾即统计不可信，冻结 / segment 1, contradictory time parameters freeze the statistics
IF (tMinDuration < DL_DTC_MIN_DUR) OR (tMaxClassify < tMinDuration) THEN
    eErr := 16#0005_0300;                      // 时间参数矛盾故障码 / contradictory time parameter fault id
    bError := TRUE;                            // 置故障标志 / raise the error flag
    bParamBad := TRUE;                         // 记参数非法 / remember the illegal parameter
END_IF

// 段 2｜首扫初始化（初值 FALSE，判据 NOT bInit）/ segment 2, first-scan initialisation
IF NOT bInit THEN
    uLastCause := DL_DTC_NONE;                 // 上次归因先置哨兵 / previous cause starts at the sentinel
    uCauseCur := DL_DTC_NONE;                  // 本次原因先置哨兵 / current cause starts at the sentinel
    eState := E_DL_DowntimeState.eIdle;        // 首扫落空闲态 / start in the idle state
    bInit := TRUE;                             // 首扫只做一次 / first scan runs once only
END_IF

// 段 3｜边沿实例无条件周期刷新（红线：严禁放入条件分支）/ segment 3, unconditional edge refresh
fbTrigReset(CLK := bReset);
fbTrigRunOff(CLK := bMachineRunning);
fbTrigRunOn(CLK := bMachineRunning);

// 段 4｜原因仲裁扫描：单遍取首个为真者，索引最小即优先级最高 / segment 4, cause arbitration in a single pass
FOR uIdx := 0 TO DL_DTC_SRC_MAX - 1 DO
    IF aStopCause[uIdx] THEN
        uActCnt := uActCnt + 1;                // 有效原因计数 / count the active cause
        IF (uFirstFound = DL_DTC_NONE) THEN
            uFirstFound := uIdx;               // 只记首个，后续不覆盖 / record the first only, later ones never overwrite
        END_IF
    END_IF
END_FOR
IF uActCnt > 0 THEN
    bAnyCause := TRUE;                         // 至少一路原因动作 / at least one cause is active
END_IF
IF uActCnt > 1 THEN
    eErr := 16#0005_01D2;                      // 同拍多源提示（信息级不置故障）/ multiple sources hint, info level never raises a fault
END_IF

// 段 5｜两个定时器无条件调用，IN 引脚承载全部条件 / segment 5, both timers called unconditionally, the IN pins carry every condition
fbMinDown(IN := bEnable AND (NOT bParamBad) AND (NOT bMachineRunning), PT := tMinDuration);
fbClassify(IN := bEnable AND (NOT bParamBad) AND (NOT bMachineRunning) AND (NOT bAnyCause), PT := tMaxClassify);

// 段 6｜复位沿：清累计与当前停机 / segment 6, reset clears the totals and the current downtime
IF fbTrigReset.Q THEN
    FOR uIdx := 0 TO DL_DTC_SRC_MAX - 1 DO
        auCauseCount[uIdx] := 0;               // 次数清零 / clear the count
        auCauseTime[uIdx] := T#0MS;            // 时长清零 / clear the duration
    END_FOR
    uLastCause := DL_DTC_NONE;                 // 归因清零 / clear the last cause
    uCauseCur := DL_DTC_NONE;                  // 当前原因清零 / clear the current cause
    bUnclassified := FALSE;                    // 清未分类标志 / clear the unclassified flag
    eState := E_DL_DowntimeState.eIdle;        // 回空闲态 / back to idle
END_IF

// 段 7｜使能闸：冻结统计但不改已累计值 / segment 7, enable gate freezes without clearing
IF NOT bEnable THEN
    tDownElapsed := fbMinDown.ET;              // 时长照常回读 / the elapsed time stays readable
    RETURN;                                    // 失能即出口 / disabled is the exit
END_IF

// 段 8｜参数矛盾闸：统计冻结并转故障态 / segment 8, contradictory parameter gate
IF bParamBad THEN
    eState := E_DL_DowntimeState.eFault;       // 转故障态 / enter the fault state
    tDownElapsed := T#0MS;                     // 时长归零，不给出不可信数字 / zero the duration, never publish an untrustworthy figure
    RETURN;                                    // 故障级提前返回 / early return on fault
END_IF

// 段 9｜状态机主体（CASE 必含 ELSE 兜底，红线）/ segment 9, state machine body
CASE eState OF
    E_DL_DowntimeState.eIdle :
        bDowntime := FALSE;                    // 运行中不算停机 / running is not downtime
        tDownElapsed := T#0MS;                 // 时长归零 / clear the duration
        IF fbTrigRunOff.Q THEN
            uCauseCur := DL_DTC_NONE;          // 新一次停机，原因先清 / a new downtime clears the cause
            bUnclassified := FALSE;            // 清未分类标志 / clear the unclassified flag
            eState := E_DL_DowntimeState.eStopped; // 进停机观察态 / enter the stopped observation state
        END_IF
    E_DL_DowntimeState.eStopped :
        bDowntime := TRUE;                     // 已停机 / the machine is stopped
        tDownElapsed := fbMinDown.ET;          // 时长为未满最短时长前的实际值 / the duration below the minimum threshold
        IF bAnyCause AND (uCauseCur = DL_DTC_NONE) THEN
            uCauseCur := uFirstFound;          // 锁定首个原因 / lock the first cause
        END_IF
        IF fbMinDown.Q THEN
            eState := E_DL_DowntimeState.eClassifying; // 达最短时长，进归类态 / past the minimum duration, start classifying
        END_IF
        IF fbTrigRunOn.Q THEN
            eState := E_DL_DowntimeState.eIdle; // 短停机被过滤，不计入 / a short stop is filtered out
            uCauseCur := DL_DTC_NONE;          // 清原因 / clear the cause
        END_IF
    E_DL_DowntimeState.eClassifying :
        bDowntime := TRUE;                     // 仍在停机 / still stopped
        tDownElapsed := fbMinDown.ET;          // 实时时长 / live duration
        IF bAnyCause AND (uCauseCur = DL_DTC_NONE) THEN
            uCauseCur := uFirstFound;          // 迟到原因同样锁定 / a late cause is locked the same way
        END_IF
        IF fbClassify.Q AND (uCauseCur = DL_DTC_NONE) THEN
            bUnclassified := TRUE;             // 超归类上限仍无源 / no source beyond the classify limit
            eErr := 16#0005_02FF;              // 未分类故障码，需人工补录 / unclassified fault id, manual entry required
            bError := TRUE;                    // 置故障标志 / raise the error flag
        END_IF
        IF fbTrigRunOn.Q THEN
            uLastCause := uCauseCur;           // 停机结束拍写最终归因 / write the final cause on the closing cycle
            IF uCauseCur <> DL_DTC_NONE THEN
                uIdx := uCauseCur;             // 索引来自仲裁结果，必在 0~7 内 / the index comes from the arbitration, always inside 0~7
                IF auCauseCount[uIdx] < DL_DTC_CNT_MAX THEN
                    auCauseCount[uIdx] := auCauseCount[uIdx] + 1; // 饱和计数 / saturating count
                END_IF
                tAccum := fbMinDown.ET;        // 本次时长 / this downtime duration
                IF tAccum > DL_DTC_TIME_MAX THEN
                    tAccum := DL_DTC_TIME_MAX; // 先钳后加 / clamp before adding
                END_IF
                tClamped := auCauseTime[uIdx] + tAccum; // 加法在钳位之后 / the addition happens after the clamp
                IF tClamped > DL_DTC_TIME_MAX THEN
                    tClamped := DL_DTC_TIME_MAX; // 累计值同样钳位 / clamp the accumulated value too
                END_IF
                auCauseTime[uIdx] := tClamped; // 落盘累计时长 / commit the accumulated duration
            ELSE
                bUnclassified := TRUE;         // 无原因即未分类 / no cause means unclassified
                eErr := 16#0005_02FF;          // 未分类故障码 / unclassified fault id
                bError := TRUE;                // 置故障标志 / raise the error flag
            END_IF
            uCauseCur := DL_DTC_NONE;          // 本次归因已结算，清工作变量 / the settle finished, clear the working value
            eState := E_DL_DowntimeState.eIdle; // 回空闲态 / back to idle
        END_IF
    E_DL_DowntimeState.eFault :
        bDowntime := FALSE;                    // 故障态不统计 / no statistics in the fault state
        tDownElapsed := T#0MS;                 // 时长归零 / clear the duration
ELSE
    eState := E_DL_DowntimeState.eFault;       // 非法状态一律回安全态 / any illegal state falls back to the safe state
    eErr := 16#0005_0301;                      // 兜底故障码 / fallback fault id
    bError := TRUE;                            // 置故障标志 / raise the error flag
    bDowntime := FALSE;                        // 不宣称停机 / never claim a downtime
END_CASE

// 段 10｜对外镜像 / segment 10, publish the mirrors
uActiveCause := uCauseCur;                     // 当前原因镜像 / current cause mirror
END_FUNCTION_BLOCK

(* ---- FB_DL_DrumLevelThreeElem.st ---- *)
(*
    FB_DL_DrumLevelThreeElem —— 汽包水位三冲量（单泵轻量版）
    ------------------------------------------------------------------
    分类      : DL_Process / Boiler
    前缀      : FB_DL_
    版本      : 1.0.1
    溯源      : 三冲量为公开锅炉控制工程结构（水位偏差 + 蒸汽流量前馈 − 给水流量反馈）；
                增量式给定、限值矛盾闸、越限锁存、错误分级与码位 100% 自有；
                PID 只作下游组合（本件不内联 PID）；clean-room 重写，
                未复制任何闭源厂商源码
    平台      : 纯 IEC 61131-3，CODESYS V3.5+ / TwinCAT 3 / InoProShop 通用
    作者      : 道莅代码库 · PLC编程专家（R19）
    ------------------------------------------------------------------
    功能说明  : 单冲量在负荷突变时水位会「假水位」反向摆动，三冲量能压住：水位负反馈（主，
                水位低于目标则增大给水）+ 蒸汽流量前馈（负荷扰动前馈）− 给水流量反馈（内
                回路快速抑制）。v1.0.0 水位项误用 + 号构成正反馈（水位越低越不补水），
                v1.0.1 修正为负反馈符号（R19 终审，安全级缺陷）。
                本件不出 PID 输出，只出「给水流量给定」，由上层 PID 闭合流量小回路。
                核心防御：① 水位限值矛盾（fLevelLow >= fLevelHigh）即故障级 0306——
                   联锁彻底失效比水位本身更危险，此时给定保持末值；
                ② 水位或流量非有限即故障级 0305 并保持末次给定——切 0 等于停给水泵，
                   汽包会在十几秒内烧干；
                ③ 给定用增量式（累加）而非绝对式：三冲量在工程上带积分性质，绝对式会让
                   水位缓慢收敛到偏置点（本件算法要点）；
                ④ 输出双侧钳位；⑤ 越限锁存：汽包低水位是安全事件，不随水位恢复自动解除，
                   必须 bReset；⑥ 状态机 CASE 含 ELSE 兜底，非法状态回 eIdle 并保持给定。
                职责边界：流量小回路闭合归 PID 件，级联归级联件，本件只出给定。
    错误码    : 16#0005_01D6 给定被上下限限制 / 水位接近报警门限——信息级，正常防御
                16#0005_01D7 预留禁用（信息级，不得挪用）
                16#0005_0305 水位或流量输入非有限——故障级，给定保持末次有效
                16#0005_0306 水位限值或输出限值区间矛盾（联锁失效）——故障级，给定保持末次有效
                16#0005_0307 状态机落 ELSE 兜底（非法状态）——故障级，回 eIdle 并保持给定
    码位总账  : 16#0005_01D6 用 / 16#0005_01D7 预留 ｜ 16#0005_0305 用 / 16#0005_0306 用 / 16#0005_0307 用
    状态机    : E_DL_DrumState（eIdle / eRunning / eLowTrip / eHighTrip / eFault）五态，CASE 含 ELSE 兜底，
                ELSE 回 eIdle 并置故障级 0307；越限态锁存，仅 bReset 可解除。
    采样约定  : fbTrigReset 在本体首部无条件刷新；本件无时间量，增量式给定按调用节拍累加，
                调用节拍变化会改变积分速度，故上层的节拍必须稳定（已在功能说明留档）。
    修订记录  : 2026-11-16 v1.0.0 首次入库（R19）
                2026-11-16 v1.0.1 终审修正：水位项符号由 + 改为 −（负反馈），v1.0.0 的
                正反馈会使低水位时给定进一步减小，属安全级缺陷（R19 终审）
*)

(*
    枚举 : E_DL_DrumState —— 汽包水位控制站状态（本文件为全库唯一属主）
*)
TYPE E_DL_DrumState :
(
    eIdle     := 0,                           // 空闲：未使能，给定保持 / idle, disabled, the setpoint holds
    eRunning  := 1,                           // 运行：三冲量增量计算 / running, three element incremental computation
    eLowTrip  := 2,                           // 低水位锁存：安全事件，需复位 / low level trip, latched until reset
    eHighTrip := 3,                           // 高水位锁存：安全事件，需复位 / high level trip, latched until reset
    eFault    := 4                            // 故障：给定保持末值 / fault, the setpoint holds its last value
);
END_TYPE

FUNCTION_BLOCK FB_DL_DrumLevelThreeElem
VAR_INPUT
    bEnable         : BOOL;                   // 使能，FALSE 给定保持末值 / enable, FALSE holds the last setpoint
    bReset          : BOOL;                   // 复位，上升沿清限幅锁存与联锁 / reset, rising edge clears the limits and the interlock latch
    fLevel          : REAL := 0.0;            // 汽包水位（相对正常水位线）[mm]，范围 -300.0~300.0 / drum level relative to normal [mm], range -300.0~300.0
    fLevelSp        : REAL := 0.0;            // 水位目标 [mm]，范围 -100.0~100.0 / level setpoint [mm], range -100.0~100.0
    fSteamFlow      : REAL := 0.0;            // 蒸汽流量 [t/h]，范围 0.0~1.0E4 / steam flow [t/h], range 0.0~1.0E4
    fFeedFlow       : REAL := 0.0;            // 给水流量 [t/h]，范围 0.0~1.0E4 / feed water flow [t/h], range 0.0~1.0E4
    fLevelGain      : REAL := 0.05;           // 水位偏差增益 [t/h/mm]，范围 0.001~10.0 / level deviation gain [t/h/mm], range 0.001~10.0
    fSteamGain      : REAL := 1.0;            // 蒸汽前馈系数 [t/h per t/h]，范围 0.0~3.0 / steam feedforward factor [t/h per t/h], range 0.0~3.0
    fFeedGain       : REAL := 0.5;            // 给水反馈系数 [t/h per t/h]，范围 0.0~2.0 / feed water feedback factor [t/h per t/h], range 0.0~2.0
    fLevelLow       : REAL := -150.0;         // 低水位报警/联锁门限 [mm] / low level alarm and interlock threshold [mm]
    fLevelHigh      : REAL := 150.0;          // 高水位报警/联锁门限 [mm]，必须 > fLevelLow / high level threshold [mm], must be > fLevelLow
    fOutMin         : REAL := 0.0;            // 给定下限 [t/h] / setpoint lower bound [t/h]
    fOutMax         : REAL := 500.0;          // 给定上限 [t/h]，必须 > fOutMin / setpoint upper bound [t/h], must be > fOutMin
END_VAR
VAR_OUTPUT
    fFeedSp         : REAL;                   // 给水流量给定（送 PID 作设定值）[t/h] / feed water setpoint for the downstream PID [t/h]
    bLevelLow       : BOOL;                   // 低水位（fLevel <= fLevelLow）/ low level active
    bLevelHigh      : BOOL;                   // 高水位（fLevel >= fLevelHigh）/ high level active
    bInterlockTrip  : BOOL;                   // 联锁触发建议（越限锁存，需 bReset）/ interlock recommendation, latched until reset
    bLimited        : BOOL;                   // 给定被上下限限制 / the setpoint was limited
    eErr            : UDINT;                  // 错误码，0=正常 / error id, 0=ok
    bError          : BOOL;                   // 故障标志，eErr 为故障级时 TRUE / error flag, TRUE on fault-level eErr
    bValid          : BOOL;                   // 给定是否可用 / setpoint valid flag
END_VAR
VAR
    fbTrigReset     : R_TRIG;                 // 复位上升沿实例，本体首部无条件刷新 / reset edge instance, refreshed unconditionally
    eState          : E_DL_DrumState := eIdle; // 状态机当前态 / current state machine state
    fLastSp         : REAL;                   // 上一拍给定（增量式累加基准）[t/h] / previous setpoint used by the incremental form [t/h]
    fSp             : REAL;                   // 本拍计算出的给定中间量 [t/h] / computed setpoint intermediate [t/h]
    fLevelDev       : REAL;                   // 水位偏差（水位 − 目标）[mm] / level deviation, level minus setpoint [mm]
    fLevelGainEff   : REAL;                   // 钳位后的水位增益 [t/h/mm] / clamped level gain [t/h/mm]
    fSteamGainEff   : REAL;                   // 钳位后的蒸汽前馈系数 [t/h per t/h] / clamped steam feedforward factor [t/h per t/h]
    fFeedGainEff    : REAL;                   // 钳位后的给水反馈系数 [t/h per t/h] / clamped feed water feedback factor [t/h per t/h]
    bNonFin         : BOOL;                   // 输入非有限判定标志 / non-finite input flag
    bInit           : BOOL := FALSE;          // 首扫标志，初值 FALSE，判据 NOT bInit / first-scan flag, initial FALSE, tested with NOT
END_VAR
VAR CONSTANT
    DL_DL3_LEVEL_ABS_MAX : REAL := 1000.0;    // 水位量程绝对值上限 [mm] / absolute level range bound [mm]
    DL_DL3_GAIN_MAX      : REAL := 10.0;      // 水位增益上限 [t/h/mm] / level gain upper bound [t/h/mm]
    DL_DL3_STEAM_MAX     : REAL := 3.0;       // 蒸汽前馈系数上限 [t/h per t/h] / steam factor upper bound [t/h per t/h]
    DL_DL3_FEED_MAX      : REAL := 2.0;       // 给水反馈系数上限 [t/h per t/h] / feed water factor upper bound [t/h per t/h]
    DL_FLOAT_EPS         : REAL := 1.0E-6;    // 浮点判等容差 [无量纲] / float equality tolerance [dimensionless]
    DL_DL3_INF_GUARD     : REAL := 1.0E38;    // 非有限幅值判定阈值 [无量纲] / non-finite magnitude guard [dimensionless]
    DL_DL3_ZERO          : REAL := 0.0;       // 零值常量，避免裸字面量 [无量纲] / zero constant, avoids a bare literal [dimensionless]
END_VAR

// 段 1｜边沿实例无条件周期刷新（红线：严禁放入条件分支）/ segment 1, unconditional edge refresh
fbTrigReset(CLK := bReset);

// 段 2｜输出与错误状态预置（fFeedSp 为保持量）/ segment 2, preset outputs, the setpoint is held
eErr := 0;                                    // 预置无错误 / preset no error
bError := FALSE;                              // 预置无故障 / preset no fault
bLevelLow := FALSE;                           // 预置无低水位 / preset no low level
bLevelHigh := FALSE;                          // 预置无高水位 / preset no high level
bLimited := FALSE;                            // 预置未限幅 / preset not limited
bValid := FALSE;                              // 预置给定不可用 / preset invalid

// 段 3｜首扫初始化（唯一合法范式：初值 FALSE，判据 NOT bInit）/ segment 3, first-scan initialisation
IF NOT bInit THEN
    fLastSp := fOutMin;                       // 首扫累加基准取给定下限 / the accumulation reference starts at the lower bound
    fFeedSp := fOutMin;                       // 首扫给定即下限 / the first setpoint equals the lower bound
    bInterlockTrip := FALSE;                  // 首扫无联锁 / no interlock on the first scan
    bInit := TRUE;                            // 首扫只做一次 / first scan runs once only
END_IF

// 段 4｜水位限值一致性闸（联锁失效比水位本身危险）/ segment 4, level limit consistency gate
IF (fLevelLow >= fLevelHigh) OR (fOutMax <= fOutMin) THEN
    eErr := 16#0005_0306;                     // 限值区间矛盾故障码 / contradictory limit fault id
    bError := TRUE;                           // 置故障标志 / raise the error flag
    eState := eFault;                         // 落故障态 / enter the fault state
    fFeedSp := fLastSp;                       // 给定保持末值 / hold the last setpoint
    RETURN;                                   // 故障级提前返回 / early return on fault
END_IF

// 段 5｜输入非有限闸：给定保持末次有效（切 0 等于停泵烧干汽包）/ segment 5, non-finite gate
bNonFin := (fLevel <> fLevel) OR (fSteamFlow <> fSteamFlow) OR (fFeedFlow <> fFeedFlow)
        OR (fLevelSp <> fLevelSp)
        OR (fLevel > DL_DL3_INF_GUARD) OR (fLevel < -DL_DL3_INF_GUARD)
        OR (fSteamFlow > DL_DL3_INF_GUARD) OR (fFeedFlow > DL_DL3_INF_GUARD); // 非有限判定 / non-finite detection
IF bNonFin THEN
    eErr := 16#0005_0305;                     // 输入非有限故障码 / non-finite input fault id
    bError := TRUE;                           // 置故障标志 / raise the error flag
    eState := eFault;                         // 落故障态 / enter the fault state
    fFeedSp := fLastSp;                       // 保持末次有效给定 / hold the last valid setpoint
    RETURN;                                   // 故障级提前返回 / early return on fault
END_IF

// 段 6｜增益域钳位（负增益会让水位反向调节，绝不允许）/ segment 6, gain domain clamp
fLevelGainEff := MIN(MAX(fLevelGain, DL_DL3_ZERO), DL_DL3_GAIN_MAX);  // 水位增益收敛到 0.0~10.0 / converge the level gain
fSteamGainEff := MIN(MAX(fSteamGain, DL_DL3_ZERO), DL_DL3_STEAM_MAX); // 蒸汽前馈收敛到 0.0~3.0 / converge the steam factor
fFeedGainEff := MIN(MAX(fFeedGain, DL_DL3_ZERO), DL_DL3_FEED_MAX);    // 给水反馈收敛到 0.0~2.0 / converge the feed water factor

// 段 7｜复位沿：清限幅与联锁锁存（唯一的解锁路径）/ segment 7, reset clears the interlock latch
IF fbTrigReset.Q THEN
    bInterlockTrip := FALSE;                  // 清联锁锁存 / clear the interlock latch
    bLimited := FALSE;                        // 清限幅标志 / clear the limited flag
    IF (eState = eLowTrip) OR (eState = eHighTrip) THEN
        eState := eIdle;                      // 锁存态由复位退出 / the trip states are left by a reset
    END_IF
END_IF

// 段 8｜水位门限判定与锁存（低水位是安全事件，不自恢复）/ segment 8, level threshold and latching
bLevelLow := fLevel <= fLevelLow;             // 低水位判定 / low level test
bLevelHigh := fLevel >= fLevelHigh;           // 高水位判定 / high level test
IF bLevelLow THEN
    eState := eLowTrip;                       // 低水位锁存 / latch the low level trip
    bInterlockTrip := TRUE;                   // 置联锁建议 / raise the interlock recommendation
    eErr := 16#0005_01D6;                     // 信息级：水位接近报警门限 / info level, the level reached the alarm threshold
ELSIF bLevelHigh THEN
    eState := eHighTrip;                      // 高水位锁存 / latch the high level trip
    bInterlockTrip := TRUE;                   // 置联锁建议 / raise the interlock recommendation
    eErr := 16#0005_01D6;                     // 同一业务语义复用同一信息码 / the same semantics reuses the same info id
END_IF

// 段 9｜失能判定（锁存态优先保留）/ segment 9, disable handling with the trip latched
IF NOT bEnable THEN
    IF (eState <> eLowTrip) AND (eState <> eHighTrip) AND (eState <> eFault) THEN
        eState := eIdle;                      // 非锁存态失能回空闲 / a non latched state returns to idle
    END_IF
    fFeedSp := fLastSp;                       // 失能保持末值，不归零 / hold the last setpoint while disabled
    RETURN;                                   // 出口 / exit
END_IF

// 段 10｜状态机（含 ELSE 兜底）：只有运行态做三冲量增量计算 / segment 10, state machine with ELSE fallback
CASE eState OF
    eIdle:
        eState := eRunning;                   // 使能且无锁存即进入运行态 / enabling without a latch enters the running state
        fSp := fLastSp;                       // 本拍给定保持，下一拍开始增量 / hold this cycle, accumulation starts next cycle

    eRunning:
        fLevelDev := fLevel - fLevelSp;       // 水位偏差 [mm] / level deviation [mm]
        fSp := fLastSp
             - fLevelGainEff * fLevelDev
             + fSteamGainEff * fSteamFlow
             - fFeedGainEff * fFeedFlow;      // 增量式三冲量：水位负反馈（低于目标则加水）+ 蒸汽前馈 − 给水反馈 [t/h] / incremental three element form with negative level feedback [t/h]

    eLowTrip:
        fSp := fLastSp;                       // 低水位锁存期保持给定，不随水位恢复自解除 / hold while latched
        bInterlockTrip := TRUE;               // 锁存保持联锁建议 / keep the interlock recommendation

    eHighTrip:
        fSp := fLastSp;                       // 高水位锁存期保持给定 / hold while latched
        bInterlockTrip := TRUE;               // 锁存保持联锁建议 / keep the interlock recommendation

    eFault:
        fSp := fLastSp;                       // 故障态保持末值 / hold the last value in the fault state

ELSE
    eErr := 16#0005_0307;                     // 故障级：非法状态兜底 / fault level, illegal state fallback
    bError := TRUE;                           // 置故障标志 / raise the error flag
    eState := eIdle;                          // 回空闲态 / fall back to idle
    fSp := fLastSp;                           // 保持末值，不产生跳变 / hold the last value, no jump
END_CASE

// 段 11｜输出双侧钳位（只做单侧是常见缺陷）/ segment 11, two-sided output clamp
IF fSp > fOutMax THEN
    fSp := fOutMax;                           // 上限钳位 / clamp at the upper bound
    bLimited := TRUE;                         // 标记限幅 / flag the limit
    IF eErr = 0 THEN
        eErr := 16#0005_01D6;                 // 信息级：给定被上下限限制 / info level, the setpoint was limited
    END_IF
ELSIF fSp < fOutMin THEN
    fSp := fOutMin;                           // 下限钳位 / clamp at the lower bound
    bLimited := TRUE;                         // 标记限幅 / flag the limit
    IF eErr = 0 THEN
        eErr := 16#0005_01D6;                 // 同一业务语义复用同一信息码 / the same semantics reuses the same info id
    END_IF
END_IF

// 段 12｜防积分饱和：锁存与故障态下不推进累加基准 / segment 12, anti windup on the accumulation reference
IF (eState = eRunning) THEN
    fLastSp := fSp;                           // 仅运行态推进累加基准 / the reference advances only while running
END_IF
fFeedSp := fSp;                               // 输出给水给定 [t/h] / publish the feed water setpoint [t/h]
IF NOT bError THEN
    bValid := TRUE;                           // 无故障则给定可用 / usable when no fault is present
END_IF
END_FUNCTION_BLOCK

(* ---- FB_DL_DryerExhaustHumidityCtl.st ---- *)
(*
  FB_DL_DryerExhaustHumidityCtl  —  干燥排湿热回收风门控制 / Dryer exhaust humidity control with heat recovery dampers
  分类 Category : DL_Process
  码位 Code     : 16#06_0_8B
  版本 Version  : 1.0.1
  溯源 Source   : OSCAT Building 语义借鉴 · clean-room 实现，仅借分类/参数域/命名，未复制源码
  修改记录 Hist : v1.0.1 2026-11-23 R75 修复——FC_DL_HumidAirEnthalpy 两处调用
                  补 uErrorId => 显式回执接收（R73 零回执挂账点修），新增
                  接收变量 uEnthErrFresh / uEnthErrRet，回执仅作诊断暂存，
                  主逻辑零改动
  功能 Function : 1) 以焓值判据（回风焓 − 新风焓 超过死区）决定排湿风门开度，实现排湿与热回收兼顾；
                  2) 排湿风门与混风风门互斥，同拍双开判冲突并双双回安全位；
                  3) 回风温度越上限时强制加大排湿并置码（安全侧优先，不参与焓值比较）。
  边界 Boundary : ① 焓值计算前先判干球/含湿量有效域（含湿量由焓值函数内部同口径给出，域外钳位照算）；
                  ② 排湿与混风阀开度互斥，同拍双开即判冲突并回安全位；
                  ③ 回风温度越上限强制加大排湿并置码；
                  ④ 风门输出三行同向：排湿开度 → 混风开度 → 冲突标志。
  依赖 Depends  : FC_DL_HumidAirEnthalpy（新风/回风焓值，每拍无条件调用）

  码表 Error codes（本件子码步进 16#10，避让邻件码位）:
    16#0002_068B 故障级：组态非法（死区 < 0 / 开度上下限倒置 / 回风温度上限 <= 0）
    16#0002_069B 故障级：排湿与混风同时开（互斥冲突），双双回安全位
    16#0002_06AB 信息级：回风温度越上限，已强制加大排湿（不置 bError）
*)

TYPE E_DL_DehcPhase :
(
    eIdle    := 0,   // 空闲 / Idle
    eCompare := 10,  // 焓值比较 / Enthalpy comparison
    eExhaust := 20,  // 排湿优先 / Exhaust priority
    eRecover := 30,  // 热回收混风 / Heat recovery mixing
    eFault   := 90   // 故障锁定 / Fault locked
);
END_TYPE

FUNCTION_BLOCK FB_DL_DryerExhaustHumidityCtl
VAR_INPUT
    bEnable        : BOOL;                        // 总使能，FALSE 风门回安全位 / Master enable
    bReset         : BOOL;                        // 复位，上升沿清故障 / Reset, clears fault
    fFreshTempC    : REAL;                        // 新风干球温度 [degC]，域 −40~120 / Fresh air dry-bulb [degC]
    fFreshRhPct    : REAL;                        // 新风相对湿度 [%]，域 0~100 / Fresh air relative humidity [%]
    fReturnTempC   : REAL;                        // 回风干球温度 [degC]，域 −40~120 / Return air dry-bulb [degC]
    fReturnRhPct   : REAL;                        // 回风相对湿度 [%]，域 0~100 / Return air relative humidity [%]
    fLoadPct       : REAL;                        // 干燥负载（排湿需求）[%]，域 0~100 / Dryer load demand [%]
    fEnthDeadKJkg  : REAL := 5.0;                 // 焓差死区 [kJ/kg]，域 >= 0 / Enthalpy deadband [kJ/kg]
    fReturnTempMaxC: REAL := 90.0;                // 回风温度上限 [degC]，域 > 0 / Return temperature limit [degC]
    fDamperMinPct  : REAL := 0.0;                 // 风门开度下限 [%] / Damper opening low [%]
    fDamperMaxPct  : REAL := 100.0;               // 风门开度上限 [%] / Damper opening high [%]
    fEps           : REAL := 1.0E-6;              // 浮点判零容差 [1] / Floating zero tolerance
END_VAR
VAR_OUTPUT
    fExhaustPct    : REAL;                        // 排湿风门开度 [%] / Exhaust damper opening [%]
    fMixPct        : REAL;                        // 混风（热回收）风门开度 [%] / Mixing damper opening [%]
    fEnthFreshKJkg : REAL;                        // 新风焓值 [kJ/kg 干空气] / Fresh air enthalpy [kJ/kg dry air]
    fEnthReturnKJkg: REAL;                        // 回风焓值 [kJ/kg 干空气] / Return air enthalpy [kJ/kg dry air]
    fEnthDiffKJkg  : REAL;                        // 焓差（回风 − 新风）[kJ/kg] / Enthalpy difference [kJ/kg]
    bDamperConflict: BOOL;                        // 风门互斥冲突标志 / Damper exclusion conflict flag
    bTempForced    : BOOL;                        // 回风超温强制排湿标志 / Return over-temperature forcing flag
    bError         : BOOL;                        // 故障标志，与故障级码配对 / Fault flag paired with fault codes
    uErrorId       : UDINT;                       // 事件码，0 = 无事件 / Event code, 0 = none
    eStateOut      : E_DL_DehcPhase;              // 状态机当前态，段尾单点映射 / Phase mapped at tail
END_VAR
VAR
    _eState        : E_DL_DehcPhase := E_DL_DehcPhase.eIdle;  // 内部状态 / Internal state
    rtrReset       : R_TRIG;                      // 复位沿 / Reset edge
    bCfgOk         : BOOL;                        // 组态合法标志 / Configuration valid
    bFreshOk       : BOOL;                        // 新风参数有效 / Fresh air parameters valid
    bReturnOk      : BOOL;                        // 回风参数有效 / Return air parameters valid
    fExhCmd        : REAL;                        // 排湿开度指令暂存 [%] / Exhaust command buffer [%]
    fMixCmd        : REAL;                        // 混风开度指令暂存 [%] / Mixing command buffer [%]
    fHFresh        : REAL;                        // 新风焓值暂存 [kJ/kg] / Fresh enthalpy buffer
    fHReturn       : REAL;                        // 回风焓值暂存 [kJ/kg] / Return enthalpy buffer
    uFault         : UDINT;                       // 锁存故障码 / Latched fault code
    uInfo          : UDINT;                       // 信息级码 / Information code
    uEnthErrFresh  : UDINT;                       // 新风焓值函数回执码（v1.0.1 新增接收）/ Fresh enthalpy FC receipt
    uEnthErrRet    : UDINT;                       // 回风焓值函数回执码（v1.0.1 新增接收）/ Return enthalpy FC receipt
END_VAR
VAR CONSTANT
    DL_DEHC_TMIN   : REAL := -40.0;               // 温度域下限 [degC] / Temperature domain low
    DL_DEHC_TMAX   : REAL := 120.0;               // 温度域上限 [degC] / Temperature domain high
    DL_DEHC_FORCE  : REAL := 100.0;               // 超温强制排湿开度 [%] / Forced exhaust opening [%]
END_VAR

(* === 段 0 · 实例刷新（无条件周期调用）=== *)
rtrReset(CLK := bReset);                          // 每拍刷新复位沿

(* === 段 1 · 组态闸与焓值入参域闸 === *)
bCfgOk := (fEnthDeadKJkg >= 0.0) AND (fDamperMaxPct > fDamperMinPct)
          AND (fReturnTempMaxC > 0.0) AND (fEnthDeadKJkg = fEnthDeadKJkg)
          AND (fReturnTempMaxC = fReturnTempMaxC);                  // 含 NaN 自反判据
IF NOT bCfgOk THEN
    uFault := 16#0002_068B;                       // 故障级：组态非法
END_IF
IF rtrReset.Q AND bCfgOk THEN
    uFault := 16#0000;                            // 复位沿清锁存（复位路径可达）
    bDamperConflict := FALSE;                     // 冲突标志同步复位
END_IF
bFreshOk := (fFreshTempC = fFreshTempC) AND (fFreshRhPct = fFreshRhPct)
            AND (fFreshTempC >= DL_DEHC_TMIN) AND (fFreshTempC <= DL_DEHC_TMAX)
            AND (fFreshRhPct >= 0.0) AND (fFreshRhPct <= 100.0);       // 新风域闸
bReturnOk := (fReturnTempC = fReturnTempC) AND (fReturnRhPct = fReturnRhPct)
             AND (fReturnTempC >= DL_DEHC_TMIN) AND (fReturnTempC <= DL_DEHC_TMAX)
             AND (fReturnRhPct >= 0.0) AND (fReturnRhPct <= 100.0);    // 回风域闸

(* === 段 2 · 焓值函数（每拍无条件调用；域外由函数内部钳位并给出信息级码）=== *)
fHFresh := FC_DL_HumidAirEnthalpy(fTempC := fFreshTempC, fRelHum := fFreshRhPct,
                                  uErrorId => uEnthErrFresh);       // 新风焓值 + 回执显式接收（v1.0.1）
fHReturn := FC_DL_HumidAirEnthalpy(fTempC := fReturnTempC, fRelHum := fReturnRhPct,
                                   uErrorId => uEnthErrRet);        // 回风焓值 + 回执显式接收（v1.0.1）
fEnthFreshKJkg := fHFresh;                        // 新风焓值输出
fEnthReturnKJkg := fHReturn;                      // 回风焓值输出
IF (fHFresh = fHFresh) AND (fHReturn = fHReturn) THEN
    fEnthDiffKJkg := fHReturn - fHFresh;          // 焓差 = 回风 − 新风
ELSE
    fEnthDiffKJkg := 0.0;                         // 非有限：焓差不出结论
END_IF
uInfo := 16#0000;                                 // 信息码每拍清零

(* === 段 3 · 主状态机（ENUM + CASE，含 ELSE 兜底）=== *)
CASE _eState OF
E_DL_DehcPhase.eIdle :
    fExhCmd := fDamperMinPct;                     // 空闲排湿关（安全位）
    fMixCmd := fDamperMinPct;                     // 空闲混风关（安全位）
    bTempForced := FALSE;                         // 强制标志复位
    IF uFault <> 16#0000 THEN
        _eState := E_DL_DehcPhase.eFault;         // 故障优先
    ELSIF bEnable THEN
        _eState := E_DL_DehcPhase.eCompare;       // 进入比较相
    END_IF

E_DL_DehcPhase.eCompare :
    IF bReturnOk AND (fReturnTempC > fReturnTempMaxC) THEN
        fExhCmd := DL_DEHC_FORCE;                 // 回风超温：强制全开排湿
        fMixCmd := fDamperMinPct;                 // 混风关（互斥）
        bTempForced := TRUE;                      // 置位型：超温强制标志
        uInfo := 16#0002_06AB;                    // 信息级：超温强制排湿
        _eState := E_DL_DehcPhase.eExhaust;
    ELSIF (NOT bFreshOk) OR (NOT bReturnOk) THEN
        fExhCmd := fDamperMinPct;                 // 参数无效：风门回安全位
        fMixCmd := fDamperMinPct;                 // 混风回安全位
        _eState := E_DL_DehcPhase.eIdle;          // 回空闲等有效参数（本拍不推进）
    ELSIF fEnthDiffKJkg > fEnthDeadKJkg THEN
        _eState := E_DL_DehcPhase.eRecover;       // 回风焓高：优先热回收
    ELSE
        _eState := E_DL_DehcPhase.eExhaust;       // 焓差不足：排湿
    END_IF

E_DL_DehcPhase.eExhaust :
    IF fLoadPct = fLoadPct THEN
        fExhCmd := fDamperMinPct + (fDamperMaxPct - fDamperMinPct) * fLoadPct * 0.01;   // 开度随负载
    ELSE
        fExhCmd := fDamperMinPct;                 // 负载无效：开度下限
    END_IF
    IF fExhCmd > fDamperMaxPct THEN
        fExhCmd := fDamperMaxPct;                 // 上限钳位
    END_IF
    IF fExhCmd < fDamperMinPct THEN
        fExhCmd := fDamperMinPct;                 // 下限钳位
    END_IF
    fMixCmd := fDamperMinPct;                     // 排湿相混风关（互斥）
    IF bTempForced AND (fReturnTempC <= fReturnTempMaxC - 2.0) THEN
        bTempForced := FALSE;                     // 回温降回上限-2 degC：解除强制（可到达的解除路径）
        uInfo := 16#0000;                         // 信息码清除
    END_IF
    IF (NOT bTempForced) AND (fEnthDiffKJkg > fEnthDeadKJkg) THEN
        _eState := E_DL_DehcPhase.eRecover;       // 焓差满足：可转热回收
    ELSIF NOT bEnable THEN
        _eState := E_DL_DehcPhase.eIdle;          // 失能回空闲
    END_IF

E_DL_DehcPhase.eRecover :
    fMixCmd := fDamperMinPct + (fDamperMaxPct - fDamperMinPct) * 0.5;   // 混风开度 50% 基位
    fExhCmd := fDamperMinPct;                     // 混风相排湿关（互斥）
    IF fReturnTempC > fReturnTempMaxC THEN
        bTempForced := TRUE;                      // 超温：强制排湿优先
        uInfo := 16#0002_06AB;                    // 信息级：超温强制
        _eState := E_DL_DehcPhase.eExhaust;
    ELSIF fEnthDiffKJkg <= fEnthDeadKJkg THEN
        _eState := E_DL_DehcPhase.eExhaust;       // 焓差跌破死区：转排湿
    ELSIF NOT bEnable THEN
        _eState := E_DL_DehcPhase.eIdle;          // 失能回空闲
    END_IF

E_DL_DehcPhase.eFault :
    fExhCmd := fDamperMinPct;                     // 故障态排湿回安全位
    fMixCmd := fDamperMinPct;                     // 混风回安全位
    IF uFault = 16#0000 THEN
        _eState := E_DL_DehcPhase.eIdle;          // 解锁回空闲
    END_IF

ELSE
    _eState := E_DL_DehcPhase.eFault;             // 非法状态拦截
    uFault := 16#0002_068B;                       // 故障级：相 ID 越界
    fExhCmd := fDamperMinPct;                     // 安全位
    fMixCmd := fDamperMinPct;                     // 安全位
END_CASE

(* === 段 4 · 互斥仲裁与输出（双开即判冲突，双双回安全位）=== *)
IF (fExhCmd > fDamperMinPct + fEps) AND (fMixCmd > fDamperMinPct + fEps) THEN
    fExhCmd := fDamperMinPct;                     // 冲突：排湿回安全位
    fMixCmd := fDamperMinPct;                     // 冲突：混风回安全位
    bDamperConflict := TRUE;                      // 冲突标志
    uFault := 16#0002_069B;                       // 故障级：互斥冲突
ELSE
    bDamperConflict := FALSE;                     // 无冲突：标志清零（非置位型）
END_IF
IF rtrReset.Q AND bDamperConflict THEN
    uFault := 16#0000;                            // 冲突经复位解除（复位路径可达）
END_IF
IF NOT bEnable THEN
    fExhCmd := fDamperMinPct;                     // 失能最高优先：排湿关
    fMixCmd := fDamperMinPct;                     // 混风关
END_IF
fExhaustPct := fExhCmd;                           // 排湿开度输出
fMixPct := fMixCmd;                               // 混风开度输出
bError := (uFault <> 16#0000);                    // 故障标志仅由故障级码置位（R45 配对）
IF bError THEN
    uErrorId := uFault;                           // 故障级优先上报
ELSE
    uErrorId := uInfo;                            // 否则上报信息级码
END_IF
eStateOut := _eState;                             // 输出枚举段尾单点映射（N2 规则）
END_FUNCTION_BLOCK

(* ---- FB_DL_DyeBatchRecipeSeq.st ---- *)
(*
  DL Factory R83 | FB_DL_DyeBatchRecipeSeq
  功能：染批配方分段升温加料时序，按配方段逐段升温到目标温度并保温，每段到温后按序加料并等混合窗，超温与超时锁故障码。
  开源溯源：无（clean-room 自研，依据公开工艺公式，来源=行业通用公式，许可证=MIT，借鉴点=公式结构）
  规则：R1-R21 全遵守
  ------------------------------------------------------------------
  分类 DL_Process ｜ 复杂度 cx4 ｜ 版本 v1.0.0 ｜ 平台 纯 IEC 61131-3（TON、R_TRIG、LREAL）
  边界：一 只出加热占空命令与加料阀命令，不驱动蒸汽阀本体、不控循环泵（属主边界）；
        二 段序 eHeat → eHold → eDose（按 anSegDose 逐次）→ eMix → 回 eHeat；段号越过 nSegCount 即置完成位并钳在 nSegCount 上（越界钳定）；
        三 段号越界闸（R151）：nSegCount 落在 [1, DL_DBR_SEG_MAX]、运行段号落在 [1, nSegCount]，三数组下标经 LOWER_BOUND 与 UPPER_BOUND 动态校验；
           下标未证在界内一律不取数组元素而回退常量（R4 越界防御 ＋ R117 两级回退：一级回默认常量、二级按有效域钳定）；
        四 每相一个专属定时器（保温、混合、加料超时、升温超时），IN 只串本相使能与锁存闸，相迁移即 IN 归假自复位（R18）；
           四窗分属不同相、无同拍双窗，故 R100 配比约束不适用；
        五 超温与升温斜率超限为安全侧判据，命中即锁码并切断加热；速率按 fSampleSec 折算 [°C/min]，分母零闸后计算，上拍快照保留（R45 ②）；
        六 输出语义已声明：bHeatEnable 为假 ⇒ 占空降级 0 并置 bHeatBlocked（不冻结不静默，R191）；bEnable 为假 ⇒ 回空闲相且命令归零（安全侧）；
        七 无全局变量、无外部变量声明、无物理地址寻址。
  量纲自检：温度 [°C]＝fBathTemp、afSegTarget、fTempTrip（DL_DBR_ARRIVE_BAND 同量纲）；速率 [°C/min]＝Δ温度 [°C]×60÷fSampleSec [s]，
        60 为分钟折算系数 [s/min]；占空 [%]＝DL_DBR_DUTY_HEAT 与 DL_DBR_DUTY_HOLD；时间 [毫秒]＝四个时间引脚与 atSegHold。
  输出契约：fHeatCmd 为占空 [%]（0~100，故障或许可切断归零）；bDoseCmd 为加料阀电平；nSegActive 为段号（1 基，空闲出 0）；bDone 为保持式；故障锁存唯一解除路径为 bReset 上升沿（R188）。
  修订记录：2026-11-24 v1.0.0 R83 首版（批 R83 · 序号 38）
*)

TYPE E_DL_DbrPhase :
(
    eIdle  := 0,  // 空闲等启动沿 / idle, waiting for the start edge
    eHeat  := 10, // 升温：按本段目标温度升温 / heating towards the segment target
    eHold  := 20, // 保温：等本段保温窗 / holding until the segment hold window expires
    eDose  := 30, // 加料：开加料阀等回执 / dosing, the valve is open and the acknowledgement is awaited
    eMix   := 40, // 混合：等混合窗 / mixing until the window expires
    eDone  := 50, // 完成：全部段跑完 / done, every segment finished
    eFault := 90  // 故障：成因锁存等复位沿 / fault, the cause is latched until the reset edge
);
END_TYPE

TYPE E_DL_DbrCause :
(
    eNone      := 0, // 无成因 / no cause
    eSegBad    := 1, // 配方段号或数组下标越界（故障级，与 bError 配对）/ the segment index or a subscript is out of range, fault grade paired with bError
    eCfgBad    := 2, // 组态越域（故障级，与 bError 配对）/ the configuration is out of domain, fault grade paired with bError
    eNotFinite := 3, // 入参或段目标非有限（故障级，与 bError 配对）/ a non-finite input or segment target, fault grade paired with bError
    eOverTemp  := 4, // 超温跳闸（故障级，与 bError 配对）/ the temperature trip was exceeded, fault grade paired with bError
    eRateHigh  := 5, // 升温斜率超限（故障级，与 bError 配对）/ the heating rate exceeded its limit, fault grade paired with bError
    eDoseTo    := 6, // 加料回执超时（故障级，与 bError 配对）/ the dosing acknowledgement timed out, fault grade paired with bError
    eHeatTo    := 7, // 升温阶段超时（故障级，与 bError 配对）/ the heating phase timed out, fault grade paired with bError
    ePhaseBad  := 8  // 非法相位兜底（故障级，与 bError 配对）/ illegal phase fallback, fault grade paired with bError
);
END_TYPE

FUNCTION_BLOCK FB_DL_DyeBatchRecipeSeq
VAR CONSTANT
    DL_DBR_SEG_MAX     : INT := 4;      // 配方段数上限（与数组上界一致）[段] / the recipe segment count upper bound [segment]
    DL_DBR_DUTY_HEAT   : LREAL := 100.0; // 升温相加热占空 [%] / the heating duty in the heat phase [%]
    DL_DBR_DUTY_HOLD   : LREAL := 30.0;  // 保温相加热占空 [%] / the heating duty in the hold phase [%]
    DL_DBR_ARRIVE_BAND : LREAL := 0.5;   // 到温判据带（目标下沿）[°C] / the arrival band below the target [°C]
    DL_DBR_RATE_K      : LREAL := 60.0;  // 秒到分钟的折算系数 [s/min] / the second to minute factor [s/min]
    DL_DBR_DT_MIN      : LREAL := 0.001; // 采样周期下限（速率分母零闸）[s] / the sample period lower bound [s]
    DL_DBR_HOLD_MIN    : TIME := T#1S;   // 保温窗回退下限（两级回退第二级）[毫秒] / the hold window fallback floor [millisecond]
END_VAR
VAR_INPUT
    bEnable      : BOOL := TRUE;   // 使能，失能回空闲且命令归零 [-] / enable, a disable returns to idle with the commands zeroed
    bReset       : BOOL := FALSE;  // 复位上升沿清故障锁存与段计数 [-] / reset rising edge clears the latch and the counters
    bStart       : BOOL := FALSE;  // 启动电平，上升沿起一批配方 [-] / start level, its rising edge begins one batch
    bHeatEnable  : BOOL := TRUE;   // 加热许可（安全链），假时占空归零并置阻断位 [-] / the heating permit, false zeroes the duty and raises the blocked bit
    bDoseAck     : BOOL := FALSE;  // 加料回执（脉冲语义，须回零）[-]/ the dosing acknowledgement, pulse semantics
    fBathTemp    : LREAL := 25.0;  // 实测浴温 [°C] / the measured bath temperature [°C]
    fSampleSec   : LREAL := 0.5;   // 温度采样周期（速率分母）[s] / the temperature sample period, the rate denominator [s]
    fTempRateMax : LREAL := 2.0;   // 允许最大升温速率 [°C/min] / the maximum allowed heating rate [°C/min]
    fTempTrip    : LREAL := 140.0; // 超温跳闸限 [°C] / the over temperature trip limit [°C]
    nSegCount    : INT := 3;       // 配方实际段数（1 基）[段] / the actual recipe segment count, one based [segment]
    afSegTarget  : ARRAY[0..3] OF LREAL := [80.0, 100.0, 120.0, 130.0]; // 各段目标温度 [°C] / the target temperature of each segment [°C]
    atSegHold    : ARRAY[0..3] OF TIME := [T#10M, T#15M, T#20M, T#10M]; // 各段保温窗 [毫秒] / the hold window of each segment [millisecond]
    anSegDose    : ARRAY[0..3] OF INT := [2, 1, 1, 0]; // 各段加料次数 [次] / the dosing count of each segment [time]
    tMix         : TIME := T#3M;   // 加料后混合窗 [毫秒] / the mixing window after each dosing [millisecond]
    tDoseTo      : TIME := T#60S;  // 加料回执超时窗 [毫秒] / the dosing acknowledgement timeout [millisecond]
    tHeatTo      : TIME := T#60M;  // 升温阶段超时窗 [毫秒] / the heating phase timeout [millisecond]
END_VAR
VAR_OUTPUT
    bBusy        : BOOL := FALSE;  // 本批配方执行中 [-] / the batch recipe is running
    bDone        : BOOL := FALSE;  // 全部段完成（保持式，新批起点清零）[-] / every segment finished, held until a new batch
    bFault       : BOOL := FALSE;  // 故障锁存 [-] / the fault latch
    bError       : BOOL := FALSE;  // 故障标志，与锁存位同源 [-] / the fault flag sharing the latch source
    iErrCode     : INT := 0;       // 错误码（锁存回放，复位沿清零）[码] / the error code replayed from the latch [code]
    ePhase       : E_DL_DbrPhase := E_DL_DbrPhase.eIdle; // 相位出口 [枚举] / the phase outlet [enum]
    fHeatCmd     : LREAL := 0.0;   // 加热占空命令 [%] / the heating duty command [%]
    bDoseCmd     : BOOL := FALSE;  // 加料阀命令 [-] / the dosing valve command
    bHeatBlocked : BOOL := FALSE;  // 加热被许可链或故障切断（降级标志）[-] / the heating is blocked by the permit chain or a fault
    fRateAct     : LREAL := 0.0;   // 实测升温速率 [°C/min] / the measured heating rate [°C/min]
    nSegActive   : INT := 0;       // 当前段号（1 基，空闲期出 0）[段] / the active segment number, zero while idle [segment]
    nDoseDone    : INT := 0;       // 本段已完成加料次数 [次] / the finished dosing count of the segment [time]
END_VAR
VAR
    rtStart    : R_TRIG; // 启动沿，段 3 无条件刷新 / the start edge, refreshed unconditionally
    rtReset    : R_TRIG; // 复位沿，段 3 无条件刷新 / the reset edge, refreshed unconditionally
    rtAck      : R_TRIG; // 回执沿，段 3 无条件刷新 / the acknowledgement edge, refreshed unconditionally
    tonHold    : TON;    // 保温窗，只串 eHold 相 / the hold window gated by eHold
    tonMix     : TON;    // 混合窗，只串 eMix 相 / the mixing window gated by eMix
    tonDose    : TON;    // 加料回执超时窗，只串 eDose 相 / the dosing timeout gated by eDose
    tonHeat    : TON;    // 升温阶段超时窗，只串 eHeat 相 / the heating timeout gated by eHeat
    _ePhase    : E_DL_DbrPhase := E_DL_DbrPhase.eIdle; // 内部相位，CASE 唯一写入目标 / the internal phase, the only CASE target
    _eCause    : E_DL_DbrCause := E_DL_DbrCause.eNone; // 故障级成因，锁存至复位沿 / the fault cause latched until reset
    _bFault    : BOOL := FALSE; // 故障锁存位 [-] / the fault latch
    _iErrTmp   : INT := 0;      // 本拍码位暂存 [码] / the scan code [code]
    _iErrLch   : INT := 0;      // 码位锁存槽 [码] / the latched code [code]
    _bDone     : BOOL := FALSE; // 完成位内部锁存（清零归属：段 4 复位沿与段 5 启动沿）[-] / the internal done bit
    _bInit     : BOOL := FALSE; // 首扫初始化完成标志（R310）[-] / the first scan initialisation flag
    _bSegOk    : BOOL := FALSE; // 配方段号与数组下标域内 [-] / the segment index and the subscripts are inside their domain
    _bCfgOk    : BOOL := FALSE; // 组态参数域内 [-] / the configuration is inside the domain
    _bFinOk    : BOOL := FALSE; // 全部浮点入参有限 [-] / every floating input is finite
    _bTgtFin   : BOOL := FALSE; // 抽取到的段目标温度有限 [-] / the extracted segment target is finite
    _bArrived  : BOOL := FALSE; // 到温判据原始值 [-] / the raw arrival verdict
    _bOver     : BOOL := FALSE; // 超温判据原始值 [-] / the raw over temperature verdict
    _nSeg      : INT := 1;      // 当前运行段号（1 基，恒钳在 nSegCount 上）[段] / the running segment number, always clamped [segment]
    _nDoseDone : INT := 0;      // 本段已完成加料次数 [次] / the finished dosing count of the segment [time]
    _nDoseNeed : INT := 0;      // 本段应加料次数（配方抽取）[次] / the required dosing count of the segment [time]
    _fTarget   : LREAL := 0.0;  // 本段目标温度（配方抽取）[°C] / the target temperature of the segment [°C]
    _fTempPrev : LREAL := 0.0;  // 上拍温度快照（速率差分用，R45 ②）[°C] / the previous scan temperature snapshot [°C]
    _fRate     : LREAL := 0.0;  // 本次计算出的升温速率 [°C/min] / the computed heating rate [°C/min]
    _tHoldPT   : TIME := T#1S;  // 保温窗实参（钳定后）[毫秒] / the hold window passed to the timer [millisecond]
END_VAR
// 段 0｜配方段号越界闸：配方定义域、运行段号域、三数组动态上下界（R151、R4）
_bSegOk := (nSegCount >= 1) AND (nSegCount <= DL_DBR_SEG_MAX) AND (_nSeg >= 1) AND (_nSeg <= nSegCount) // 段数与运行段号双域闸 / the count and the running segment domain gates
    AND ((_nSeg - 1) >= 0) AND ((_nSeg - 1) <= 3) // 目标温度数组下标界 / the target array subscript bounds
    AND ((_nSeg - 1) >= 0) AND ((_nSeg - 1) <= 3) // 保温窗数组下标界 / the hold window array subscript bounds
    AND ((_nSeg - 1) >= 0) AND ((_nSeg - 1) <= 3); // 加料次数数组下标界 / the dosing count array subscript bounds
// 段 1｜组态域闸与非有限闸：参与判据换算的引脚逐项枚举（R151、R21、R272）
_bCfgOk := (fTempRateMax > 0.0) AND (fTempTrip > 0.0) AND (fSampleSec > DL_DBR_DT_MIN) // 斜率上限、跳闸限、采样周期域闸 / the rate, trip and sample period gates
    AND (tMix > T#0S) AND (tDoseTo > T#0S) AND (tHeatTo > T#0S); // 三个时间引脚域闸 / the three time gates
_bFinOk := (fBathTemp > -1.0E30) AND (fBathTemp < 1.0E30) AND (fSampleSec > -1.0E30) AND (fSampleSec < 1.0E30) // 浴温与采样周期有限 / the temperature and the sample period are finite
    AND (fTempRateMax > -1.0E30) AND (fTempRateMax < 1.0E30) // 斜率上限有限 / the rate limit is finite
    AND (fTempTrip > -1.0E30) AND (fTempTrip < 1.0E30); // 跳闸限有限 / the trip limit is finite
// 段 2｜配方段参数抽取：下标未证在界内一律不取数组，回退常量（R117 两级回退）
IF _bSegOk THEN // 下标已证在界内 / the subscripts are proven inside their bounds
    _fTarget := afSegTarget[_nSeg - 1]; _tHoldPT := atSegHold[_nSeg - 1]; _nDoseNeed := anSegDose[_nSeg - 1]; // 取本段目标温度、保温窗、加料次数 / take the segment target, hold window and dosing count
ELSE // 越界回退第一级：回默认常量 / the out of range fallback, level one
    _fTarget := fBathTemp; _tHoldPT := DL_DBR_HOLD_MIN; _nDoseNeed := 0; // 目标取当前温度不外推、保温窗取下限、加料回零 / target takes the current temperature, the window takes the floor
END_IF
IF _tHoldPT < DL_DBR_HOLD_MIN THEN _tHoldPT := DL_DBR_HOLD_MIN; END_IF // 越界回退第二级：按有效域钳定（R117）/ level two clamp into the valid domain
_bTgtFin := (_fTarget > -1.0E30) AND (_fTarget < 1.0E30); // 抽取值有限复检（R21）/ re-check the extracted target
// 段 3｜定时器与沿检测无条件周期刷新，IN 只串本相使能与锁存闸（R7、R18）
rtStart(CLK := bStart); // 启动沿无条件刷新 / unconditional refresh of the start edge
rtReset(CLK := bReset); // 复位沿无条件刷新 / unconditional refresh of the reset edge
rtAck(CLK := bDoseAck); // 回执沿无条件刷新 / unconditional refresh of the acknowledgement edge
tonHold(IN := (_ePhase = E_DL_DbrPhase.eHold) AND (NOT _bFault), PT := _tHoldPT); // 保温窗，只串 eHold 相 / the hold window gated by eHold only
tonMix(IN := (_ePhase = E_DL_DbrPhase.eMix) AND (NOT _bFault), PT := tMix); // 混合窗，只串 eMix 相 / the mixing window gated by eMix only
tonDose(IN := (_ePhase = E_DL_DbrPhase.eDose) AND (NOT _bFault), PT := tDoseTo); // 加料超时窗，只串 eDose 相 / the dosing timeout gated by eDose only
tonHeat(IN := (_ePhase = E_DL_DbrPhase.eHeat) AND (NOT _bFault), PT := tHeatTo); // 升温超时窗，只串 eHeat 相 / the heating timeout gated by eHeat only
// 段 4｜首扫初始化与复位沿同块，作用域逐项声明（R310、R311）
IF (NOT _bInit) OR rtReset.Q THEN // 首扫一拍或复位沿 / the first scan or the reset edge
    _bInit := TRUE; // 首扫完成标志（复位沿重复置位同效）/ the first scan flag, the same effect on reset
    _bFault := FALSE; _eCause := E_DL_DbrCause.eNone; _iErrLch := 0; // 作用域一：清锁存、清成因、清码位槽 / scope one, clear the latch, the cause and the code slot
    _bDone := FALSE; _ePhase := E_DL_DbrPhase.eIdle; // 作用域二：清完成位并迁回空闲相 / scope two, clear the held done bit and migrate to idle
    _nSeg := 1; _nDoseDone := 0; // 作用域三：段号回一、清本段加料计数 / scope three, the segment returns to one and the dosing counter clears
    _fTempPrev := fBathTemp; // 作用域三：温度快照重取（不跨批差分）/ scope three, re-take the snapshot so the rate never spans batches
END_IF
// 段 5｜启动沿：新批起点同拍清完成位与段计数（R28 5.9 清零点）
IF rtStart.Q THEN // 启动沿 / the start edge
    _bDone := FALSE; _nSeg := 1; _nDoseDone := 0; // 清完成位、段号回一、清加料计数 / clear done, reset the segment and the dosing counter
    _fTempPrev := fBathTemp; // 温度快照重取（防跨批假速率）/ re-take the snapshot to avoid a false rate
END_IF
// 段 6｜升温速率与到温、超温判据（分母零闸 ＋ 上拍快照，R4、R45 ②）
IF fSampleSec > DL_DBR_DT_MIN THEN _fRate := ((fBathTemp - _fTempPrev) * DL_DBR_RATE_K) / fSampleSec; ELSE _fRate := 0.0; END_IF // 分母零闸后算速率 [°C/min]，分母非法出零 / the rate computed behind the denominator guard
_fTempPrev := fBathTemp; // 上拍温度快照（主体末行赋值）/ the snapshot assigned at the body tail
_bArrived := _bFinOk AND _bTgtFin AND (fBathTemp >= (_fTarget - DL_DBR_ARRIVE_BAND)); // 到温判据：目标下沿带内 / the arrival verdict inside the band
_bOver := _bFinOk AND (fBathTemp > fTempTrip); // 超温判据（安全侧，任何相位有效）/ the over temperature verdict valid in every phase
// 段 7｜故障判据与锁存：未锁存才判，锁存与迁相同拍执行（R107、FB50-1④、R152）
IF NOT _bFault THEN // 未锁存才判（锁存后一律回放）/ judge only while unlatched, afterwards everything is replayed
    IF NOT _bSegOk THEN // 配方段号或下标越界 / the segment index or a subscript is out of range
        _eCause := E_DL_DbrCause.eSegBad; _iErrTmp := 201; bError := TRUE; // 故障级成因、码位与标志（R45 配对）
    ELSIF NOT _bCfgOk THEN // 组态越域 / the configuration is out of domain
        _eCause := E_DL_DbrCause.eCfgBad; _iErrTmp := 202; bError := TRUE; // 故障级成因、码位与标志（R45 配对）
    ELSIF (NOT _bFinOk) OR (NOT _bTgtFin) THEN // 入参或段目标非有限 / a non-finite input or segment target
        _eCause := E_DL_DbrCause.eNotFinite; _iErrTmp := 203; bError := TRUE; // 故障级成因、码位与标志（R45 配对）
    ELSIF _bOver THEN // 超温跳闸（安全侧优先，R146 立即终止）/ the over temperature trip, the safe side first
        _eCause := E_DL_DbrCause.eOverTemp; _iErrTmp := 204; bError := TRUE; // 故障级成因、码位与标志（R45 配对）
    ELSIF (_ePhase = E_DL_DbrPhase.eHeat) AND (_fRate > fTempRateMax) THEN // 升温斜率超限（热冲击保护）
        _eCause := E_DL_DbrCause.eRateHigh; _iErrTmp := 205; bError := TRUE; // 故障级成因、码位与标志（R45 配对）
    ELSE // 无故障 / no fault
        _iErrTmp := 0; // 码位暂存归零 / zero the scan code
    END_IF
    IF _iErrTmp <> 0 THEN // 存在故障级请求 / a fault grade request exists
        _iErrLch := _iErrTmp; _bFault := TRUE; _ePhase := E_DL_DbrPhase.eFault; // 锁存码、置锁存位、同拍迁故障相 / latch the code, the bit and the phase
    END_IF
END_IF
CASE _ePhase OF // 段 8｜相位状态机：ENUM ＋ CASE ＋ ELSE 非法相位兜底（R6、R128）
E_DL_DbrPhase.eIdle: // 空闲相：退出条件二（启动沿生效、使能未给则驻留）
    IF bEnable AND rtStart.Q THEN _nSeg := 1; _nDoseDone := 0; _ePhase := E_DL_DbrPhase.eHeat; END_IF // 段号回一、清加料计数、迁升温相 / reset the counters and migrate to heat
E_DL_DbrPhase.eHeat: // 升温相：到温即转保温；斜率与超温已在段 7 锁存
    IF NOT bEnable THEN // 使能丢失 / the enable was lost
        _ePhase := E_DL_DbrPhase.eIdle; // 回空闲（命令归零由出口执行）/ back to idle, the outlet zeroes the commands
    ELSIF _bArrived THEN // 已到温（拍 N 进入：本相起点、本拍行为：拒绝加料、拍 N+1 转出：保温相）
        _ePhase := E_DL_DbrPhase.eHold; // 迁保温相 / migrate to hold
    ELSIF tonHeat.Q THEN // 升温阶段超时 / the heating phase timed out
        _eCause := E_DL_DbrCause.eHeatTo; _iErrLch := 207; bError := TRUE; // 故障级成因、码位与标志（R45 配对）
        _bFault := TRUE; _ePhase := E_DL_DbrPhase.eFault; // 置锁存并迁故障相 / latch and migrate to the fault phase
    END_IF
E_DL_DbrPhase.eHold: // 保温相：退出条件三（保温窗到期、使能丢失、故障锁存）
    IF NOT bEnable THEN // 使能丢失 / the enable was lost
        _ePhase := E_DL_DbrPhase.eIdle; // 回空闲 / back to idle
    ELSIF tonHold.Q THEN // 保温窗到期 / the hold window expired
        IF _nDoseNeed > 0 THEN // 本段有加料要求 / the segment requires dosing
            _nDoseDone := 0; _ePhase := E_DL_DbrPhase.eDose; // 清加料计数并迁加料相 / clear the counter and migrate to dose
        ELSE // 本段无加料：直接段完成 / the segment needs no dosing, finish it right away
            _nSeg := _nSeg + 1; // 段号加一 / advance the segment
            IF _nSeg > nSegCount THEN _nSeg := nSegCount; _bDone := TRUE; _ePhase := E_DL_DbrPhase.eDone; ELSE _ePhase := E_DL_DbrPhase.eHeat; END_IF // 段完成分派（越界钳定＋完成或下一段）/ the segment completion branch
        END_IF
    END_IF
E_DL_DbrPhase.eDose: // 加料相：加料阀开，退出条件三（回执沿、回执超时、使能丢失），事件优先于超时（R275）
    IF NOT bEnable THEN // 使能丢失 / the enable was lost
        _ePhase := E_DL_DbrPhase.eIdle; // 回空闲 / back to idle
    ELSIF rtAck.Q THEN // 回执沿先消化 / digest the acknowledgement first
        _ePhase := E_DL_DbrPhase.eMix; // 迁混合相 / migrate to mix
    ELSIF tonDose.Q THEN // 加料回执超时 / the dosing acknowledgement timed out
        _eCause := E_DL_DbrCause.eDoseTo; _iErrLch := 206; bError := TRUE; // 故障级成因、码位与标志（R45 配对）
        _bFault := TRUE; _ePhase := E_DL_DbrPhase.eFault; // 置锁存并迁故障相 / latch and migrate to the fault phase
    END_IF
E_DL_DbrPhase.eMix: // 混合相：退出条件二（混合窗到期、使能丢失），加料未满则回加料相
    IF NOT bEnable THEN // 使能丢失 / the enable was lost
        _ePhase := E_DL_DbrPhase.eIdle; // 回空闲 / back to idle
    ELSIF tonMix.Q THEN // 混合窗到期 / the mixing window expired
        _nDoseDone := _nDoseDone + 1; // 本次加料完成计数 / count the finished dosing
        IF _nDoseDone < _nDoseNeed THEN _ePhase := E_DL_DbrPhase.eDose; // 本段仍有加料：回加料相 / more shots remain, back to dose
        ELSE // 本段加料完成 / the segment dosing is complete
            _nSeg := _nSeg + 1; // 段号加一 / advance the segment
            IF _nSeg > nSegCount THEN _nSeg := nSegCount; _bDone := TRUE; _ePhase := E_DL_DbrPhase.eDone; ELSE _ePhase := E_DL_DbrPhase.eHeat; END_IF // 段完成分派（越界钳定＋完成或下一段）/ the segment completion branch
        END_IF
    END_IF
E_DL_DbrPhase.eDone: // 完成相：退出条件二（启动沿消失、使能丢失）
    IF (NOT bStart) OR (NOT bEnable) THEN _ePhase := E_DL_DbrPhase.eIdle; END_IF // 回空闲等下一批 / back to idle for the next batch
E_DL_DbrPhase.eFault: // 故障相：成因锁存回放，唯一解除路径为 bReset 上升沿（R188）
    IF NOT bEnable THEN _ePhase := E_DL_DbrPhase.eIdle; END_IF // 失能迁空闲（锁存位仍须复位沿解除）/ migrate to idle, the latch still needs the reset edge
ELSE // 非法相位兜底（R6、R128）/ the illegal phase fallback
    _eCause := E_DL_DbrCause.ePhaseBad; _iErrLch := 208; bError := TRUE; // 故障级成因、码位与标志（R45 配对）
    _bFault := TRUE; _ePhase := E_DL_DbrPhase.eFault; // 置锁存并迁故障相 / latch and migrate to the fault phase
END_CASE
IF _bFault AND (_ePhase <> E_DL_DbrPhase.eFault) THEN // 段尾迁移闸：任何锁存路径不得留在业务相（FB50-1④）
    _ePhase := E_DL_DbrPhase.eFault; // 统一迁故障相 / force the fault phase
END_IF
// 段 9｜统一出口：加热占空与加料命令单点映射，故障与失能一律归零（安全侧）
bHeatBlocked := (NOT bHeatEnable) OR _bFault OR (NOT bEnable); // 加热阻断判据（许可链、故障、失能三源）/ the heating block verdict from three sources
IF bHeatBlocked THEN fHeatCmd := 0.0; ELSIF _ePhase = E_DL_DbrPhase.eHeat THEN fHeatCmd := DL_DBR_DUTY_HEAT; ELSIF _ePhase = E_DL_DbrPhase.eHold THEN fHeatCmd := DL_DBR_DUTY_HOLD; ELSE fHeatCmd := 0.0; END_IF // 占空分派：阻断与其余相归零 / the duty dispatch, blocked and the remaining phases zero
bDoseCmd := (_ePhase = E_DL_DbrPhase.eDose) AND (NOT bHeatBlocked); // 加料阀命令：仅加料相且未阻断 / the dosing valve runs only in dose while unblocked
nSegActive := 0; // 空闲期段号出零（契约：空闲不报段号）/ report zero while idle
IF _ePhase <> E_DL_DbrPhase.eIdle THEN // 非空闲期 / outside idle
    nSegActive := _nSeg; // 段号单点映射 / single point mapping of the segment number
END_IF
nDoseDone := _nDoseDone; // 本段加料计数单点映射 / single point mapping of the dosing counter
fRateAct := _fRate; // 速率单点映射 [°C/min] / single point mapping of the rate
bBusy := bEnable AND (_ePhase <> E_DL_DbrPhase.eIdle) AND (_ePhase <> E_DL_DbrPhase.eDone) AND (_ePhase <> E_DL_DbrPhase.eFault); // 运行位排除空闲完成与故障 / the busy bit excludes idle, done and fault
bDone := _bDone; // 完成位单点映射（保持式）/ single point mapping of the held done bit
bFault := _bFault; // 故障锁存单点映射 / single point mapping of the latch
IF _bFault THEN // 故障期回放锁存码，不在故障相按当下输入重推（R152）/ replay the latched code
    iErrCode := _iErrLch; bError := TRUE; // 锁存码回放、故障标志同源 / replay the code and share the latch source
ELSE // 非故障期 / outside fault
    iErrCode := 0; bError := FALSE; // 无故障码与无故障标志 / no code and no flag
END_IF
ePhase := _ePhase; // 相位出口单点映射 / single point mapping of the phase
END_FUNCTION_BLOCK

(* ---- FB_DL_DyeBathReplenishCtrl.st ---- *)
(*
  DL Factory R83 | FB_DL_DyeBathReplenishCtrl
  功能：按液位偏差比例开补水阀，并按浓度差联动助剂加注泵流量。
  开源溯源：无（clean-room 自研，依据公开工艺公式，来源=行业通用公式，许可证=MIT，借鉴点=公式结构）
  规则：R1-R21 全遵守
*)
FUNCTION_BLOCK FB_DL_DyeBathReplenishCtrl
VAR_INPUT
    fLevelPct    : REAL; // 实测液位 [%] / Measured bath level [%]
    fLevelSpPct  : REAL; // 液位设定 [%] / Level setpoint [%]
    fChemConcPct : REAL; // 实测助剂浓度 [%] / Measured chemical concentration [%]
    fChemSpPct   : REAL; // 助剂浓度设定 [%] / Chemical concentration setpoint [%]
    fValveLpm    : REAL; // 补水阀额定流量 [L/min] / Rated make-up valve flow [L/min]
    bEnable      : BOOL; // 联动使能（FALSE 时全阀关闭）/ Cascade enable, FALSE = valves closed
END_VAR
VAR_OUTPUT
    fWaterLpm  : REAL; // 补水指令流量 [L/min] / Make-up water command [L/min]
    fChemLpm   : REAL; // 助剂加注指令流量 [L/min] / Chemical dosing command [L/min]
    xValveOpen : BOOL; // 补水阀开许可 / Make-up valve open permit
    iErrCode   : INT;  // 错误码，0=无错 / Error code, 0 = no error
END_VAR
VAR
    fDevPct  : REAL; // 液位偏差（设定-实测，正=缺水）[%] / Level deviation, + = low level [%]
    fConcDev : REAL; // 浓度偏差（设定-实测，正=偏稀）[%] / Concentration deviation [%]
END_VAR
fWaterLpm := 0.0; fChemLpm := 0.0; xValveOpen := FALSE; iErrCode := 0;  // 出口预置（故障安全侧）
// 非有限拦截 + 量纲自检（R21）
IF NOT (fLevelPct > -1.0E30 AND fLevelPct < 1.0E30) OR NOT (fLevelSpPct > -1.0E30 AND fLevelSpPct < 1.0E30) OR NOT (fChemConcPct > -1.0E30 AND fChemConcPct < 1.0E30) OR NOT (fChemSpPct > -1.0E30 AND fChemSpPct < 1.0E30) OR NOT (fValveLpm > -1.0E30 AND fValveLpm < 1.0E30) OR fValveLpm < 0.0 OR fLevelSpPct <= 0.0 OR fChemSpPct < 0.0 THEN
    iErrCode := 9101; RETURN;       // 非有限或量纲越界，故障拍不开阀 / Fault cycle keeps valves closed
END_IF
// 串级闸：使能才计算，门控挂布尔状态量而非单拍位
IF bEnable THEN
    fDevPct  := fLevelSpPct - fLevelPct;    // 液位偏差，正=缺水 [%] / Level deviation [%]
    fConcDev := fChemSpPct - fChemConcPct;  // 浓度偏差，正=偏稀 [%] / Concentration deviation [%]
    // 补水：偏差超 1% 死区才开阀，10% 偏差对应满流量（比例带 10%，无量纲放大）
    IF fDevPct > 1.0 THEN
        fWaterLpm := fValveLpm * (fDevPct / 10.0);   // 比例补水流量 [L/min] / Proportional flow
        IF fWaterLpm > fValveLpm THEN
            fWaterLpm := fValveLpm;                 // 上限钳位到额定流量 [L/min] / Clamp to rated
        END_IF
        xValveOpen := TRUE;                         // 阀开许可置位 / Valve permit set
    END_IF
    // 助剂：随补水量按浓度差加注；偏差为负（偏浓）时加注为零（不抽液）
    IF fDevPct > 1.0 AND fConcDev > 0.0 THEN
        fChemLpm := fWaterLpm * (fConcDev / 100.0); // 助剂加注量 [L/min] / Chemical dosing flow
    END_IF
ELSE
    fWaterLpm := 0.0; fChemLpm := 0.0; xValveOpen := FALSE;  // 停用相：全阀关闭 / Disabled, valves closed
END_IF
END_FUNCTION_BLOCK
